// TIA Portal project "Project2" (V17)

(* hardware
DEVICE "S7-1500/ET200MP station_1"  S7-1500 station
   slot 0: "Rail_0"  Rack  6ES7 590-1***0-0AA0
   slot 1: "PLC_2"  CPU 1515-2 PN  6ES7 515-2AM00-0AB0  V1.8
      slot 3: "CPU display_1"  6ES7591-1BA00-0AA0
      slot 32768: "PROFINET interface_1"  X1
         slot 32769: "Port_1"  X1 P1
         slot 32770: "Port_2"  X1 P2
      slot 33024: "PROFINET interface_2"  X2
         slot 33025: "Port_1"  X2 P1
*)

// ===== PLC "PLC_2"  CPU 1515-2 PN =====

// folder: UDT/S2-Process Function Unit

TYPE "UDT_IS28xx_To_Plc"
   STRUCT
      iTriggerReady : Bool;   // This bit indicates when an In-Sight device can accept a new trigger via the Trigger bit. This field is true when the Trigger Enable bit is set, and the vision system is not currently acquiring an image.
      iTriggerAck : Bool;   // This bit indicates when an In-Sight device is successfully triggered via the Trigger bit. The Trigger Acknowledge bit stays set until the Trigger bit is cleared.
      iExposureComplete : Bool;   // This bit is set when the vision system image sensor is no longer exposed to light. It is used to indicate that the part being inspected can be moved from under the vision system's field of view.
      iAcquisitionError : Bool;   // This bit is set when an In-Sight device fails to acquire an image for one of the following reasons:
      iOfflineReason_1 : Bool;   // OfflineReason_1
      iOfflineReason_2 : Bool;   // OfflineReason_2
      iOfflineReason_3 : Bool;   // OfflineReason_3
      iSystemOnline : Bool;   // This bit indicates that the In-Sight device is online and the $System.OnlineEnabled tag is True.
      iReserve_1 : Byte;   // Reserve1
      iAcquisitonID : Int;   // This ID increments on the completion of every acquisition, regardless of the trigger source, and can be used to synchronize an acquisition with its Inspection Result. The Acquisition ID is changed on the start of an acquisition. If the PLC is the trigger source, the Acquisition ID is set prior to setting the Trigger Acknowledge bit.
      iReserve_2 : Bool;   // Reserve2
      iInspectionComplete : Bool;   // This bit is toggled upon the completion of an inspection.
      iResultBufferOverRun : Bool;   // This bit is set when the Enable Results Buffer bit is set, and there are more results than the result queue can hold.
      iResultValid : Bool;   // This bit is set when the Inspected Image ID, Inspection Result Code and Inspection Results fields are valid. The bit is cleared when the Inspection Results Acknowledge bit is set.
      iCommandExecuted : Bool;   // This bit is set while a command execution is in progress.
      iCommandComplete : Bool;   // This bit is set when the command execution is completed, and cleared when the Execute Command bit has been cleare
      iCommandFailed : Bool;   // This bit is set on the completion of a command, if the command has failed to execute successfully, or if an unknown Command ID was set.
      iSetUserDataAck : Bool;   // This bit is set to acknowledge completion of the Set User Data command.
      iJobPass : Bool;   // This bit indicates the pass and/or fail state of the inspection.
      iReserve_3 : Bool;   // Reserve3
      iReserve_4 : Bool;   // Reserve4
      iReserve_5 : Bool;   // Reserve5
      iReserve_6 : Bool;   // Reserve6
      iReserve_7 : Bool;   // Reserve7
      iReserve_8 : Bool;   // Reserve8
      iError : Bool;   // This bit is set when an error has occurred, which is defined in the Error ID field.
      iErrorID : Int;   // See Error ID codes.
      iCurrentRunningJobID : Int;   // These bits indicate the pre-added number of the current job filename. A job ID is a 16 bit number from 0 to 65535, but the PLC function can only load job IDs between 0‑999.
      iCommandResultCode : Int;   // This field is used to indicate the reason a command failed to execute successfully (the code is specific to the command executed):
      iExternalSoftEventAck : Byte;   // The External Event Acknowledge will be generated after the associated script finishes its execution
      iInspectionResultData : Struct
         iInspectionID : Int;   // The acquisition ID associated with this set of results.
         iInspectionResultCode : Int;   // These bytes are used to pass the user-defined result code. The inspection result code is defined by the Result Code parameter of the WriteResultsBuffer function
         iInspectionResult : Array[1..60] of Byte;   // These bytes of the inspection tool results can be written to the currently enabled factory communication protocol via the WriteResultsBuffer function.
      END_STRUCT;
   END_STRUCT;
END_TYPE

TYPE "UDT_Plc_To_IS28xx"
   STRUCT
      qTriggerEnable : Bool;   // This field is set to enable triggering via the Trigger bit. Clear this bit to disable the network triggering mechanism
      qTrigger : Bool;   // Setting the Trigger bit will trigger an acquisition on the vision system. The Trigger Enable bit must also be set
      qClearExposureComplete : Bool;   // When this signal is held high, the Exposure Complete status will remain reset. Once this signal is set to low, the Exposure Complete status will be set to high on the next exposure completion.
      qReserve_1 : Bool;   // Reserve_1
      qReserve_2 : Bool;   // Reserve_2
      qReserve_3 : Bool;   // Reserve_3
      qReserve_4 : Bool;   // Reserve_4
      qSetOffline : Bool;   // When this bit is set, the In-Sight vision system is paused and the state of the $System.OnlineEnabledComm is false
      qBufferResultEnable : Bool;   // When this bit is set, the Inspection ID, Inspection Result and Inspection Results fields are held constant until the Inspection Results Acknowledge field has acknowledged them and been set. Up to 16 sets of results are held in the buffer. Each result must be explicitly acknowledged using the Inspection Results Acknowledge signal.
      qInspectionResultAck : Bool;   // When the Buffer Results Enable bit is set, the Inspection Results Acknowledge bit acknowledges that the PLC has received the Inspected Image ID, Inspection Result Code and Inspection Results data.
      qSetUserData : Bool;   // This bit is used to signal that new User Data is available to be read in the vision system. After latching the entire User Data area into a holding buffer, the vision system will indicate to the PLC that it has read the data, and it can start loading new data into the buffer, if required, by issuing the Set User Data Acknowledge signal.
      qExecuteCommand : Bool;   // When the Execute Command bit is set to high, the Command ID signal is read by the vision system and the associated command is executed. The signal must be held high until the Command Completed bit is set. Once the Command Completed bit is set, clearing the Execute Command bit also clears the Command Completed bit.
      qReserve_5 : Bool;   // Reserve_5
      qReserve_6 : Bool;   // Reserve_6
      qReserve_7 : Bool;   // Reserve_7
      qClearError : Bool;   // When this bit is set, it clears the Error and Error ID signals; the Clear Error bit need to be held high until the Error bit is cleared. If an error is queued, clearing this bit causes the Error and Error ID signals to be set to the next queued error code.
      qCommandID : Int;   // This field indicates the command that will be executed on the rising edge of the Execute Command bit. This signal should not be changed until the Command Completed bit has been set.
      qSoftControlInput : Byte;   // Setting the External Event allows the PLC to trigger an associated event in the Spreadsheet.
      qUserData : Array[1..60] of Byte;   // Data buffer which can be read into the spreadsheet using the ReadUserDataBuffer function. The buffer is written exactly as it appears in the PLC
   END_STRUCT;
END_TYPE

// folder: (top level)

FUNCTION_BLOCK "PR_CentreStand_Fix_Seq_V12_1026b5"   // FB1, LAD
{ S7_Optimized_Access := 'TRUE' }
VERSION : 0.1
   VAR_INPUT
      iAutoRunning : Bool;
      iFixClamp : Bool;
      iFixEmpty : Bool;
      iFixTrayPresent : Bool;
      iFixUnclamp : Bool;
      iR1DropOver : Bool;
      iR1PickOver : Bool;
      iR2OperationOver : Bool;
      iR2ServiceActivated : Bool;
      iReset_fault : Bool;
      iRobotOutofZone : Bool;
      iSstMode : Bool;
      iSstPB : Bool;
   END_VAR
   VAR_OUTPUT
      qFixClamp : Bool;
      qFixUnclamp : Bool;
      qR1ReadytoDropTray : Bool;
      qR1ReadytoPickTray : Bool;
      qR2OperationStart : Bool;
   END_VAR
   VAR_IN_OUT
      iqR2ServiceActive : Bool;
      iqR2ServiceCompleted : Bool;
   END_VAR
   VAR
      StateNo : Int;
      s138_WaitBothRbtOutAl : Bool;
      s138_WaitBothRbtOutAl_T1 : Bool;
      s138_WaitBothRbtOutAl_T2 : Bool;
      s139_FixEmpty : Bool;
      s139_FixEmpty_T1 : Bool;
      s140_FixTrayPrsntRec : Bool;
      s140_FixTrayPrsntRec_T1 : Bool;
      s140_FixTrayPrsntRec_T2 : Bool;
      s141_FixUnclampCmd : Bool;
      s141_FixUnclampCmd_T1 : Bool;
      s142_TrayRdyDropFix : Bool;
      s142_TrayRdyDropFix_T1 : Bool;
      s143_RbtDropFixChkTr : Bool;
      s143_RbtDropFixChkTr_T1 : Bool;
      s144_RbtOutAreaDrop : Bool;
      s144_RbtOutAreaDrop_T1 : Bool;
      s145_FixClamp : Bool;
      s145_FixClamp_T1 : Bool;
      s146_Rbt2AlloyOpOver : Bool;
      s146_Rbt2AlloyOpOver_T1 : Bool;
      s147_FixUnclmpCmdAft : Bool;
      s147_FixUnclmpCmdAft_T1 : Bool;
      s148_RdyPickTrayAftr : Bool;
      s148_RdyPickTrayAftr_T1 : Bool;
      s149_RbtPickTrayChkE : Bool;
      s149_RbtPickTrayChkE_T1 : Bool;
      s191_WaitRbt2OutArea : Bool;
      s191_WaitRbt2OutArea_T1 : Bool;
      sSst : Bool;
      sSstPulse : Bool;
      sSstRise : Bool;
      sStWtResetRel : Bool;
      sStWtResetRel_T1 : Bool;
   END_VAR
   VAR_TEMP
      c138_WaitBothRbtOutAl_T1 : Bool;
      c138_WaitBothRbtOutAl_T2 : Bool;
      c140_FixTrayPrsntRec_T1 : Bool;
      c140_FixTrayPrsntRec_T2 : Bool;
      tOne : Bool;
   END_VAR
   VAR_TEMP   // added for the SCL form of the ladder/FBD networks
      _w1 : Bool;
   END_VAR
BEGIN

REGION Network 1
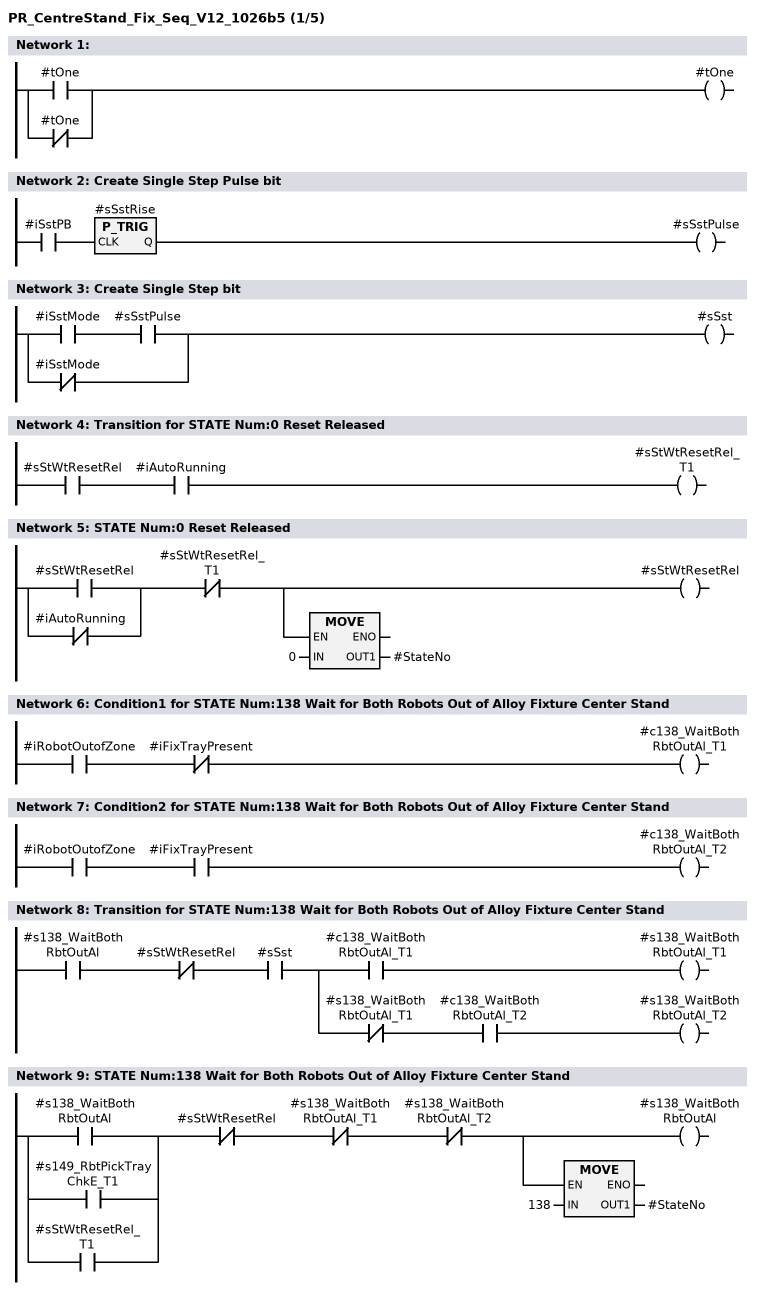
   RUNG wire#powerrail
      Contact( #tOne )
      wire#w1
      Coil( #tOne )
   END_RUNG
   RUNG wire#powerrail
      I_Contact( #tOne )
   END_RUNG wire#w1
   // the same network as SCL:
   #tOne := #tOne OR NOT #tOne;
END_REGION

REGION Network 2: Create Single Step Pulse bit
   RUNG wire#powerrail
      Contact( #iSstPB )
      P_Trig( #sSstRise )
      Coil( #sSstPulse )
   END_RUNG
   // the same network as SCL:
   #_w1 := #iSstPB AND NOT #sSstRise;   // rising edge
   #sSstRise := #iSstPB;
   #sSstPulse := #_w1;
END_REGION

REGION Network 3: Create Single Step bit
   RUNG wire#powerrail
      Contact( #iSstMode )
      Contact( #sSstPulse )
      wire#w1
      Coil( #sSst )
   END_RUNG
   RUNG wire#powerrail
      I_Contact( #iSstMode )
   END_RUNG wire#w1
   // the same network as SCL:
   #sSst := (#iSstMode AND #sSstPulse) OR NOT #iSstMode;
END_REGION

REGION Network 4: Transition for STATE Num:0 Reset Released
   RUNG wire#powerrail
      Contact( #sStWtResetRel )
      Contact( #iAutoRunning )
      Coil( #sStWtResetRel_T1 )
   END_RUNG
   // the same network as SCL:
   #sStWtResetRel_T1 := #sStWtResetRel AND #iAutoRunning;
END_REGION

REGION Network 5: STATE Num:0 Reset Released
   RUNG wire#powerrail
      Contact( #sStWtResetRel )
      wire#w1
      I_Contact( #sStWtResetRel_T1 )
      wire#w2
      Coil( #sStWtResetRel )
   END_RUNG
   RUNG wire#powerrail
      I_Contact( #iAutoRunning )
   END_RUNG wire#w1
   RUNG wire#w2
      { S7_GenerateENO := "TRUE" } Move(in := 0, out1 => #StateNo)
   END_RUNG
   // the same network as SCL:
   #sStWtResetRel := (#sStWtResetRel OR NOT #iAutoRunning) AND NOT #sStWtResetRel_T1;
   IF #sStWtResetRel THEN #StateNo := 0; END_IF;
END_REGION

REGION Network 6: Condition1 for STATE Num:138 Wait for Both Robots Out of Alloy Fixture Center Stand
   RUNG wire#powerrail
      Contact( #iRobotOutofZone )
      I_Contact( #iFixTrayPresent )
      Coil( #c138_WaitBothRbtOutAl_T1 )
   END_RUNG
   // the same network as SCL:
   #c138_WaitBothRbtOutAl_T1 := #iRobotOutofZone AND NOT #iFixTrayPresent;
END_REGION

REGION Network 7: Condition2 for STATE Num:138 Wait for Both Robots Out of Alloy Fixture Center Stand
   RUNG wire#powerrail
      Contact( #iRobotOutofZone )
      Contact( #iFixTrayPresent )
      Coil( #c138_WaitBothRbtOutAl_T2 )
   END_RUNG
   // the same network as SCL:
   #c138_WaitBothRbtOutAl_T2 := #iRobotOutofZone AND #iFixTrayPresent;
END_REGION

REGION Network 8: Transition for STATE Num:138 Wait for Both Robots Out of Alloy Fixture Center Stand
   RUNG wire#powerrail
      Contact( #s138_WaitBothRbtOutAl )
      I_Contact( #sStWtResetRel )
      Contact( #sSst )
      wire#w1
      Contact( #c138_WaitBothRbtOutAl_T1 )
      Coil( #s138_WaitBothRbtOutAl_T1 )
   END_RUNG
   RUNG wire#w1
      I_Contact( #s138_WaitBothRbtOutAl_T1 )
      Contact( #c138_WaitBothRbtOutAl_T2 )
      Coil( #s138_WaitBothRbtOutAl_T2 )
   END_RUNG
   // the same network as SCL:
   #_w1 := #s138_WaitBothRbtOutAl AND NOT #sStWtResetRel AND #sSst;
   #s138_WaitBothRbtOutAl_T1 := #_w1 AND #c138_WaitBothRbtOutAl_T1;
   #s138_WaitBothRbtOutAl_T2 := #_w1 AND NOT #s138_WaitBothRbtOutAl_T1 AND #c138_WaitBothRbtOutAl_T2;
END_REGION

REGION Network 9: STATE Num:138 Wait for Both Robots Out of Alloy Fixture Center Stand
   RUNG wire#powerrail
      Contact( #s138_WaitBothRbtOutAl )
      wire#w1
      I_Contact( #sStWtResetRel )
      I_Contact( #s138_WaitBothRbtOutAl_T1 )
      I_Contact( #s138_WaitBothRbtOutAl_T2 )
      wire#w2
      Coil( #s138_WaitBothRbtOutAl )
   END_RUNG
   RUNG wire#powerrail
      Contact( #s149_RbtPickTrayChkE_T1 )
   END_RUNG wire#w1
   RUNG wire#powerrail
      Contact( #sStWtResetRel_T1 )
   END_RUNG wire#w1
   RUNG wire#w2
      { S7_GenerateENO := "TRUE" } Move(in := 138, out1 => #StateNo)
   END_RUNG
   // the same network as SCL:
   #s138_WaitBothRbtOutAl := (#s138_WaitBothRbtOutAl OR #s149_RbtPickTrayChkE_T1 OR #sStWtResetRel_T1) AND NOT #sStWtResetRel AND NOT #s138_WaitBothRbtOutAl_T1 AND NOT #s138_WaitBothRbtOutAl_T2;
   IF #s138_WaitBothRbtOutAl THEN #StateNo := 138; END_IF;
END_REGION

REGION Network 10: Transition for STATE Num:139 Fix Empty
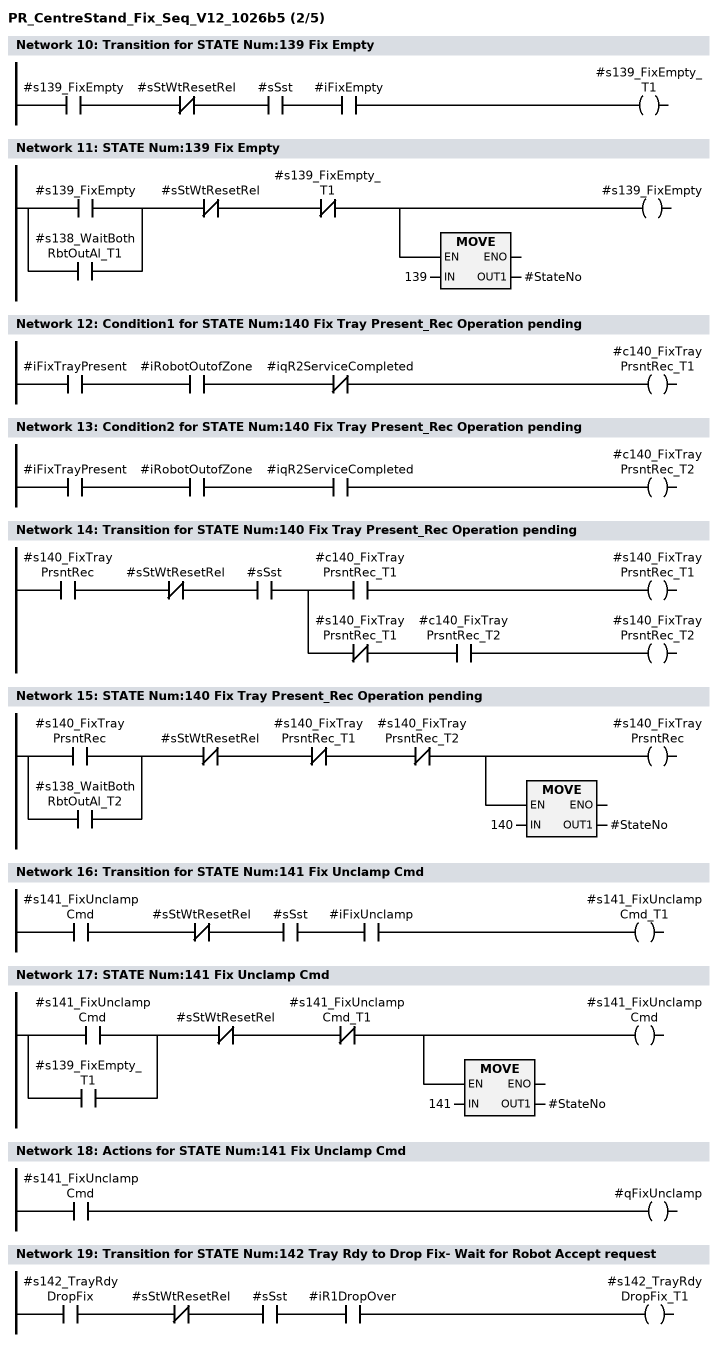
   RUNG wire#powerrail
      Contact( #s139_FixEmpty )
      I_Contact( #sStWtResetRel )
      Contact( #sSst )
      Contact( #iFixEmpty )
      Coil( #s139_FixEmpty_T1 )
   END_RUNG
   // the same network as SCL:
   #s139_FixEmpty_T1 := #s139_FixEmpty AND NOT #sStWtResetRel AND #sSst AND #iFixEmpty;
END_REGION

REGION Network 11: STATE Num:139 Fix Empty
   RUNG wire#powerrail
      Contact( #s139_FixEmpty )
      wire#w1
      I_Contact( #sStWtResetRel )
      I_Contact( #s139_FixEmpty_T1 )
      wire#w2
      Coil( #s139_FixEmpty )
   END_RUNG
   RUNG wire#powerrail
      Contact( #s138_WaitBothRbtOutAl_T1 )
   END_RUNG wire#w1
   RUNG wire#w2
      { S7_GenerateENO := "TRUE" } Move(in := 139, out1 => #StateNo)
   END_RUNG
   // the same network as SCL:
   #s139_FixEmpty := (#s139_FixEmpty OR #s138_WaitBothRbtOutAl_T1) AND NOT #sStWtResetRel AND NOT #s139_FixEmpty_T1;
   IF #s139_FixEmpty THEN #StateNo := 139; END_IF;
END_REGION

REGION Network 12: Condition1 for STATE Num:140 Fix Tray Present_Rec Operation pending
   RUNG wire#powerrail
      Contact( #iFixTrayPresent )
      Contact( #iRobotOutofZone )
      I_Contact( #iqR2ServiceCompleted )
      Coil( #c140_FixTrayPrsntRec_T1 )
   END_RUNG
   // the same network as SCL:
   #c140_FixTrayPrsntRec_T1 := #iFixTrayPresent AND #iRobotOutofZone AND NOT #iqR2ServiceCompleted;
END_REGION

REGION Network 13: Condition2 for STATE Num:140 Fix Tray Present_Rec Operation pending
   RUNG wire#powerrail
      Contact( #iFixTrayPresent )
      Contact( #iRobotOutofZone )
      Contact( #iqR2ServiceCompleted )
      Coil( #c140_FixTrayPrsntRec_T2 )
   END_RUNG
   // the same network as SCL:
   #c140_FixTrayPrsntRec_T2 := #iFixTrayPresent AND #iRobotOutofZone AND #iqR2ServiceCompleted;
END_REGION

REGION Network 14: Transition for STATE Num:140 Fix Tray Present_Rec Operation pending
   RUNG wire#powerrail
      Contact( #s140_FixTrayPrsntRec )
      I_Contact( #sStWtResetRel )
      Contact( #sSst )
      wire#w1
      Contact( #c140_FixTrayPrsntRec_T1 )
      Coil( #s140_FixTrayPrsntRec_T1 )
   END_RUNG
   RUNG wire#w1
      I_Contact( #s140_FixTrayPrsntRec_T1 )
      Contact( #c140_FixTrayPrsntRec_T2 )
      Coil( #s140_FixTrayPrsntRec_T2 )
   END_RUNG
   // the same network as SCL:
   #_w1 := #s140_FixTrayPrsntRec AND NOT #sStWtResetRel AND #sSst;
   #s140_FixTrayPrsntRec_T1 := #_w1 AND #c140_FixTrayPrsntRec_T1;
   #s140_FixTrayPrsntRec_T2 := #_w1 AND NOT #s140_FixTrayPrsntRec_T1 AND #c140_FixTrayPrsntRec_T2;
END_REGION

REGION Network 15: STATE Num:140 Fix Tray Present_Rec Operation pending
   RUNG wire#powerrail
      Contact( #s140_FixTrayPrsntRec )
      wire#w1
      I_Contact( #sStWtResetRel )
      I_Contact( #s140_FixTrayPrsntRec_T1 )
      I_Contact( #s140_FixTrayPrsntRec_T2 )
      wire#w2
      Coil( #s140_FixTrayPrsntRec )
   END_RUNG
   RUNG wire#powerrail
      Contact( #s138_WaitBothRbtOutAl_T2 )
   END_RUNG wire#w1
   RUNG wire#w2
      { S7_GenerateENO := "TRUE" } Move(in := 140, out1 => #StateNo)
   END_RUNG
   // the same network as SCL:
   #s140_FixTrayPrsntRec := (#s140_FixTrayPrsntRec OR #s138_WaitBothRbtOutAl_T2) AND NOT #sStWtResetRel AND NOT #s140_FixTrayPrsntRec_T1 AND NOT #s140_FixTrayPrsntRec_T2;
   IF #s140_FixTrayPrsntRec THEN #StateNo := 140; END_IF;
END_REGION

REGION Network 16: Transition for STATE Num:141 Fix Unclamp Cmd
   RUNG wire#powerrail
      Contact( #s141_FixUnclampCmd )
      I_Contact( #sStWtResetRel )
      Contact( #sSst )
      Contact( #iFixUnclamp )
      Coil( #s141_FixUnclampCmd_T1 )
   END_RUNG
   // the same network as SCL:
   #s141_FixUnclampCmd_T1 := #s141_FixUnclampCmd AND NOT #sStWtResetRel AND #sSst AND #iFixUnclamp;
END_REGION

REGION Network 17: STATE Num:141 Fix Unclamp Cmd
   RUNG wire#powerrail
      Contact( #s141_FixUnclampCmd )
      wire#w1
      I_Contact( #sStWtResetRel )
      I_Contact( #s141_FixUnclampCmd_T1 )
      wire#w2
      Coil( #s141_FixUnclampCmd )
   END_RUNG
   RUNG wire#powerrail
      Contact( #s139_FixEmpty_T1 )
   END_RUNG wire#w1
   RUNG wire#w2
      { S7_GenerateENO := "TRUE" } Move(in := 141, out1 => #StateNo)
   END_RUNG
   // the same network as SCL:
   #s141_FixUnclampCmd := (#s141_FixUnclampCmd OR #s139_FixEmpty_T1) AND NOT #sStWtResetRel AND NOT #s141_FixUnclampCmd_T1;
   IF #s141_FixUnclampCmd THEN #StateNo := 141; END_IF;
END_REGION

REGION Network 18: Actions for STATE Num:141 Fix Unclamp Cmd
   RUNG wire#powerrail
      Contact( #s141_FixUnclampCmd )
      Coil( #qFixUnclamp )
   END_RUNG
   // the same network as SCL:
   #qFixUnclamp := #s141_FixUnclampCmd;
END_REGION

REGION Network 19: Transition for STATE Num:142 Tray Rdy to Drop Fix- Wait for Robot Accept request
   RUNG wire#powerrail
      Contact( #s142_TrayRdyDropFix )
      I_Contact( #sStWtResetRel )
      Contact( #sSst )
      Contact( #iR1DropOver )
      Coil( #s142_TrayRdyDropFix_T1 )
   END_RUNG
   // the same network as SCL:
   #s142_TrayRdyDropFix_T1 := #s142_TrayRdyDropFix AND NOT #sStWtResetRel AND #sSst AND #iR1DropOver;
END_REGION

REGION Network 20: STATE Num:142 Tray Rdy to Drop Fix- Wait for Robot Accept request
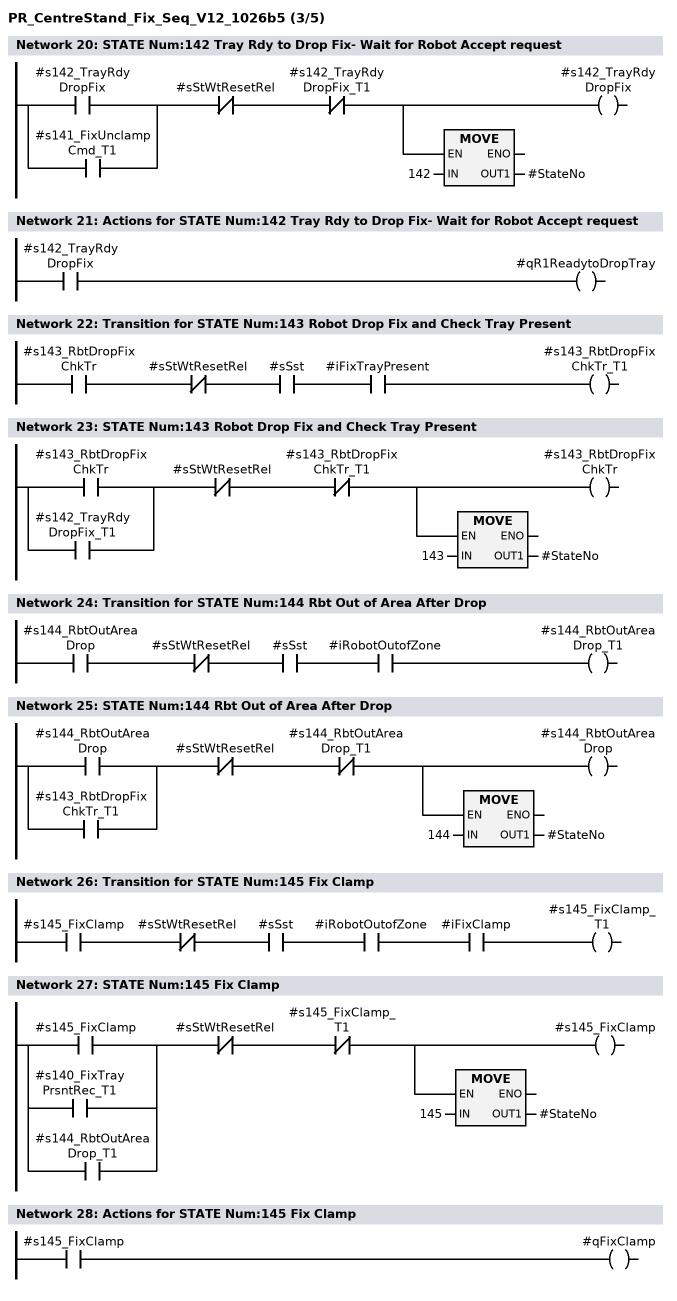
   RUNG wire#powerrail
      Contact( #s142_TrayRdyDropFix )
      wire#w1
      I_Contact( #sStWtResetRel )
      I_Contact( #s142_TrayRdyDropFix_T1 )
      wire#w2
      Coil( #s142_TrayRdyDropFix )
   END_RUNG
   RUNG wire#powerrail
      Contact( #s141_FixUnclampCmd_T1 )
   END_RUNG wire#w1
   RUNG wire#w2
      { S7_GenerateENO := "TRUE" } Move(in := 142, out1 => #StateNo)
   END_RUNG
   // the same network as SCL:
   #s142_TrayRdyDropFix := (#s142_TrayRdyDropFix OR #s141_FixUnclampCmd_T1) AND NOT #sStWtResetRel AND NOT #s142_TrayRdyDropFix_T1;
   IF #s142_TrayRdyDropFix THEN #StateNo := 142; END_IF;
END_REGION

REGION Network 21: Actions for STATE Num:142 Tray Rdy to Drop Fix- Wait for Robot Accept request
   RUNG wire#powerrail
      Contact( #s142_TrayRdyDropFix )
      Coil( #qR1ReadytoDropTray )
   END_RUNG
   // the same network as SCL:
   #qR1ReadytoDropTray := #s142_TrayRdyDropFix;
END_REGION

REGION Network 22: Transition for STATE Num:143 Robot Drop Fix and Check Tray Present
   RUNG wire#powerrail
      Contact( #s143_RbtDropFixChkTr )
      I_Contact( #sStWtResetRel )
      Contact( #sSst )
      Contact( #iFixTrayPresent )
      Coil( #s143_RbtDropFixChkTr_T1 )
   END_RUNG
   // the same network as SCL:
   #s143_RbtDropFixChkTr_T1 := #s143_RbtDropFixChkTr AND NOT #sStWtResetRel AND #sSst AND #iFixTrayPresent;
END_REGION

REGION Network 23: STATE Num:143 Robot Drop Fix and Check Tray Present
   RUNG wire#powerrail
      Contact( #s143_RbtDropFixChkTr )
      wire#w1
      I_Contact( #sStWtResetRel )
      I_Contact( #s143_RbtDropFixChkTr_T1 )
      wire#w2
      Coil( #s143_RbtDropFixChkTr )
   END_RUNG
   RUNG wire#powerrail
      Contact( #s142_TrayRdyDropFix_T1 )
   END_RUNG wire#w1
   RUNG wire#w2
      { S7_GenerateENO := "TRUE" } Move(in := 143, out1 => #StateNo)
   END_RUNG
   // the same network as SCL:
   #s143_RbtDropFixChkTr := (#s143_RbtDropFixChkTr OR #s142_TrayRdyDropFix_T1) AND NOT #sStWtResetRel AND NOT #s143_RbtDropFixChkTr_T1;
   IF #s143_RbtDropFixChkTr THEN #StateNo := 143; END_IF;
END_REGION

REGION Network 24: Transition for STATE Num:144 Rbt Out of Area After Drop
   RUNG wire#powerrail
      Contact( #s144_RbtOutAreaDrop )
      I_Contact( #sStWtResetRel )
      Contact( #sSst )
      Contact( #iRobotOutofZone )
      Coil( #s144_RbtOutAreaDrop_T1 )
   END_RUNG
   // the same network as SCL:
   #s144_RbtOutAreaDrop_T1 := #s144_RbtOutAreaDrop AND NOT #sStWtResetRel AND #sSst AND #iRobotOutofZone;
END_REGION

REGION Network 25: STATE Num:144 Rbt Out of Area After Drop
   RUNG wire#powerrail
      Contact( #s144_RbtOutAreaDrop )
      wire#w1
      I_Contact( #sStWtResetRel )
      I_Contact( #s144_RbtOutAreaDrop_T1 )
      wire#w2
      Coil( #s144_RbtOutAreaDrop )
   END_RUNG
   RUNG wire#powerrail
      Contact( #s143_RbtDropFixChkTr_T1 )
   END_RUNG wire#w1
   RUNG wire#w2
      { S7_GenerateENO := "TRUE" } Move(in := 144, out1 => #StateNo)
   END_RUNG
   // the same network as SCL:
   #s144_RbtOutAreaDrop := (#s144_RbtOutAreaDrop OR #s143_RbtDropFixChkTr_T1) AND NOT #sStWtResetRel AND NOT #s144_RbtOutAreaDrop_T1;
   IF #s144_RbtOutAreaDrop THEN #StateNo := 144; END_IF;
END_REGION

REGION Network 26: Transition for STATE Num:145 Fix Clamp
   RUNG wire#powerrail
      Contact( #s145_FixClamp )
      I_Contact( #sStWtResetRel )
      Contact( #sSst )
      Contact( #iRobotOutofZone )
      Contact( #iFixClamp )
      Coil( #s145_FixClamp_T1 )
   END_RUNG
   // the same network as SCL:
   #s145_FixClamp_T1 := #s145_FixClamp AND NOT #sStWtResetRel AND #sSst AND #iRobotOutofZone AND #iFixClamp;
END_REGION

REGION Network 27: STATE Num:145 Fix Clamp
   RUNG wire#powerrail
      Contact( #s145_FixClamp )
      wire#w1
      I_Contact( #sStWtResetRel )
      I_Contact( #s145_FixClamp_T1 )
      wire#w2
      Coil( #s145_FixClamp )
   END_RUNG
   RUNG wire#powerrail
      Contact( #s140_FixTrayPrsntRec_T1 )
   END_RUNG wire#w1
   RUNG wire#powerrail
      Contact( #s144_RbtOutAreaDrop_T1 )
   END_RUNG wire#w1
   RUNG wire#w2
      { S7_GenerateENO := "TRUE" } Move(in := 145, out1 => #StateNo)
   END_RUNG
   // the same network as SCL:
   #s145_FixClamp := (#s145_FixClamp OR #s140_FixTrayPrsntRec_T1 OR #s144_RbtOutAreaDrop_T1) AND NOT #sStWtResetRel AND NOT #s145_FixClamp_T1;
   IF #s145_FixClamp THEN #StateNo := 145; END_IF;
END_REGION

REGION Network 28: Actions for STATE Num:145 Fix Clamp
   RUNG wire#powerrail
      Contact( #s145_FixClamp )
      Coil( #qFixClamp )
   END_RUNG
   // the same network as SCL:
   #qFixClamp := #s145_FixClamp;
END_REGION

REGION Network 29: Transition for STATE Num:146 Robot-2 All Alloys Pick Or Drop Operation over
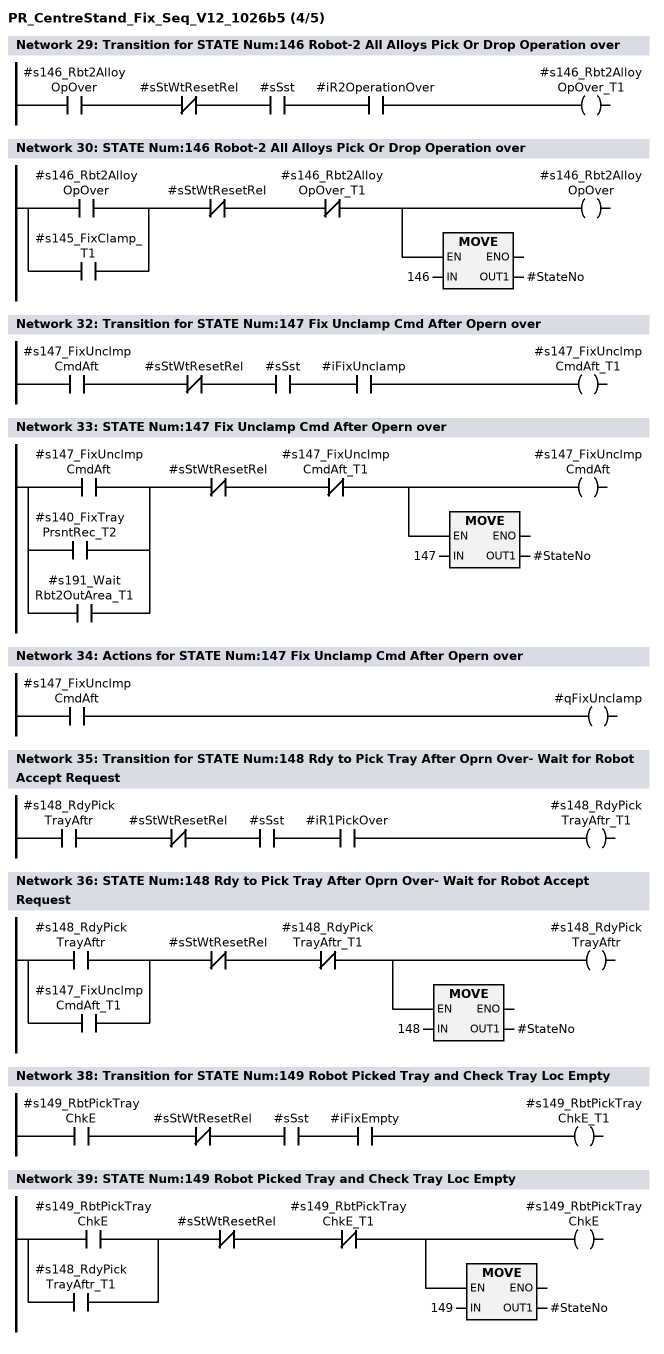
   RUNG wire#powerrail
      Contact( #s146_Rbt2AlloyOpOver )
      I_Contact( #sStWtResetRel )
      Contact( #sSst )
      Contact( #iR2OperationOver )
      Coil( #s146_Rbt2AlloyOpOver_T1 )
   END_RUNG
   // the same network as SCL:
   #s146_Rbt2AlloyOpOver_T1 := #s146_Rbt2AlloyOpOver AND NOT #sStWtResetRel AND #sSst AND #iR2OperationOver;
END_REGION

REGION Network 30: STATE Num:146 Robot-2 All Alloys Pick Or Drop Operation over
   RUNG wire#powerrail
      Contact( #s146_Rbt2AlloyOpOver )
      wire#w1
      I_Contact( #sStWtResetRel )
      I_Contact( #s146_Rbt2AlloyOpOver_T1 )
      wire#w2
      Coil( #s146_Rbt2AlloyOpOver )
   END_RUNG
   RUNG wire#powerrail
      Contact( #s145_FixClamp_T1 )
   END_RUNG wire#w1
   RUNG wire#w2
      { S7_GenerateENO := "TRUE" } Move(in := 146, out1 => #StateNo)
   END_RUNG
   // the same network as SCL:
   #s146_Rbt2AlloyOpOver := (#s146_Rbt2AlloyOpOver OR #s145_FixClamp_T1) AND NOT #sStWtResetRel AND NOT #s146_Rbt2AlloyOpOver_T1;
   IF #s146_Rbt2AlloyOpOver THEN #StateNo := 146; END_IF;
END_REGION

REGION Network 31 (STL): Actions for STATE Num:146 Robot-2 All Alloys Pick Or Drop Operation over
         A     #s146_Rbt2AlloyOpOver;
         =     #qR2OperationStart;
         A     #s146_Rbt2AlloyOpOver;
         A     #iR2ServiceActivated;
         S     #iqR2ServiceActive;
         A     #s146_Rbt2AlloyOpOver;
         A     #iR2OperationOver;
         A     #iqR2ServiceActive;
         R     #iqR2ServiceActive;
END_REGION

REGION Network 32: Transition for STATE Num:147 Fix Unclamp Cmd After Opern over
   RUNG wire#powerrail
      Contact( #s147_FixUnclmpCmdAft )
      I_Contact( #sStWtResetRel )
      Contact( #sSst )
      Contact( #iFixUnclamp )
      Coil( #s147_FixUnclmpCmdAft_T1 )
   END_RUNG
   // the same network as SCL:
   #s147_FixUnclmpCmdAft_T1 := #s147_FixUnclmpCmdAft AND NOT #sStWtResetRel AND #sSst AND #iFixUnclamp;
END_REGION

REGION Network 33: STATE Num:147 Fix Unclamp Cmd After Opern over
   RUNG wire#powerrail
      Contact( #s147_FixUnclmpCmdAft )
      wire#w1
      I_Contact( #sStWtResetRel )
      I_Contact( #s147_FixUnclmpCmdAft_T1 )
      wire#w2
      Coil( #s147_FixUnclmpCmdAft )
   END_RUNG
   RUNG wire#powerrail
      Contact( #s140_FixTrayPrsntRec_T2 )
   END_RUNG wire#w1
   RUNG wire#powerrail
      Contact( #s191_WaitRbt2OutArea_T1 )
   END_RUNG wire#w1
   RUNG wire#w2
      { S7_GenerateENO := "TRUE" } Move(in := 147, out1 => #StateNo)
   END_RUNG
   // the same network as SCL:
   #s147_FixUnclmpCmdAft := (#s147_FixUnclmpCmdAft OR #s140_FixTrayPrsntRec_T2 OR #s191_WaitRbt2OutArea_T1) AND NOT #sStWtResetRel AND NOT #s147_FixUnclmpCmdAft_T1;
   IF #s147_FixUnclmpCmdAft THEN #StateNo := 147; END_IF;
END_REGION

REGION Network 34: Actions for STATE Num:147 Fix Unclamp Cmd After Opern over
   RUNG wire#powerrail
      Contact( #s147_FixUnclmpCmdAft )
      Coil( #qFixUnclamp )
   END_RUNG
   // the same network as SCL:
   #qFixUnclamp := #s147_FixUnclmpCmdAft;
END_REGION

REGION Network 35: Transition for STATE Num:148 Rdy to Pick Tray After Oprn Over- Wait for Robot Accept Request
   RUNG wire#powerrail
      Contact( #s148_RdyPickTrayAftr )
      I_Contact( #sStWtResetRel )
      Contact( #sSst )
      Contact( #iR1PickOver )
      Coil( #s148_RdyPickTrayAftr_T1 )
   END_RUNG
   // the same network as SCL:
   #s148_RdyPickTrayAftr_T1 := #s148_RdyPickTrayAftr AND NOT #sStWtResetRel AND #sSst AND #iR1PickOver;
END_REGION

REGION Network 36: STATE Num:148 Rdy to Pick Tray After Oprn Over- Wait for Robot Accept Request
   RUNG wire#powerrail
      Contact( #s148_RdyPickTrayAftr )
      wire#w1
      I_Contact( #sStWtResetRel )
      I_Contact( #s148_RdyPickTrayAftr_T1 )
      wire#w2
      Coil( #s148_RdyPickTrayAftr )
   END_RUNG
   RUNG wire#powerrail
      Contact( #s147_FixUnclmpCmdAft_T1 )
   END_RUNG wire#w1
   RUNG wire#w2
      { S7_GenerateENO := "TRUE" } Move(in := 148, out1 => #StateNo)
   END_RUNG
   // the same network as SCL:
   #s148_RdyPickTrayAftr := (#s148_RdyPickTrayAftr OR #s147_FixUnclmpCmdAft_T1) AND NOT #sStWtResetRel AND NOT #s148_RdyPickTrayAftr_T1;
   IF #s148_RdyPickTrayAftr THEN #StateNo := 148; END_IF;
END_REGION

REGION Network 37 (STL): Actions for STATE Num:148 Rdy to Pick Tray After Oprn Over- Wait for Robot Accept Request
         A     #s148_RdyPickTrayAftr;
         =     #qR1ReadytoPickTray;
         A     #s148_RdyPickTrayAftr;
         A     #iR1PickOver;
         R     #iqR2ServiceCompleted;
END_REGION

REGION Network 38: Transition for STATE Num:149 Robot Picked Tray and Check Tray Loc Empty
   RUNG wire#powerrail
      Contact( #s149_RbtPickTrayChkE )
      I_Contact( #sStWtResetRel )
      Contact( #sSst )
      Contact( #iFixEmpty )
      Coil( #s149_RbtPickTrayChkE_T1 )
   END_RUNG
   // the same network as SCL:
   #s149_RbtPickTrayChkE_T1 := #s149_RbtPickTrayChkE AND NOT #sStWtResetRel AND #sSst AND #iFixEmpty;
END_REGION

REGION Network 39: STATE Num:149 Robot Picked Tray and Check Tray Loc Empty
   RUNG wire#powerrail
      Contact( #s149_RbtPickTrayChkE )
      wire#w1
      I_Contact( #sStWtResetRel )
      I_Contact( #s149_RbtPickTrayChkE_T1 )
      wire#w2
      Coil( #s149_RbtPickTrayChkE )
   END_RUNG
   RUNG wire#powerrail
      Contact( #s148_RdyPickTrayAftr_T1 )
   END_RUNG wire#w1
   RUNG wire#w2
      { S7_GenerateENO := "TRUE" } Move(in := 149, out1 => #StateNo)
   END_RUNG
   // the same network as SCL:
   #s149_RbtPickTrayChkE := (#s149_RbtPickTrayChkE OR #s148_RdyPickTrayAftr_T1) AND NOT #sStWtResetRel AND NOT #s149_RbtPickTrayChkE_T1;
   IF #s149_RbtPickTrayChkE THEN #StateNo := 149; END_IF;
END_REGION

REGION Network 40: Actions for STATE Num:149 Robot Picked Tray and Check Tray Loc Empty
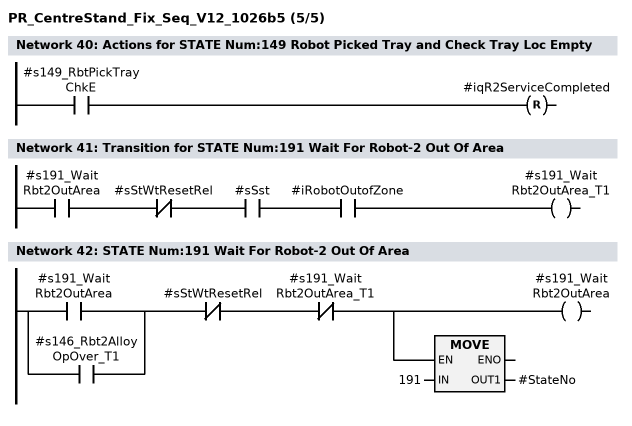
   RUNG wire#powerrail
      Contact( #s149_RbtPickTrayChkE )
      R_Coil( #iqR2ServiceCompleted )
   END_RUNG
   // the same network as SCL:
   IF #s149_RbtPickTrayChkE THEN #iqR2ServiceCompleted := FALSE; END_IF;
END_REGION

REGION Network 41: Transition for STATE Num:191 Wait For Robot-2 Out Of Area
   RUNG wire#powerrail
      Contact( #s191_WaitRbt2OutArea )
      I_Contact( #sStWtResetRel )
      Contact( #sSst )
      Contact( #iRobotOutofZone )
      Coil( #s191_WaitRbt2OutArea_T1 )
   END_RUNG
   // the same network as SCL:
   #s191_WaitRbt2OutArea_T1 := #s191_WaitRbt2OutArea AND NOT #sStWtResetRel AND #sSst AND #iRobotOutofZone;
END_REGION

REGION Network 42: STATE Num:191 Wait For Robot-2 Out Of Area
   RUNG wire#powerrail
      Contact( #s191_WaitRbt2OutArea )
      wire#w1
      I_Contact( #sStWtResetRel )
      I_Contact( #s191_WaitRbt2OutArea_T1 )
      wire#w2
      Coil( #s191_WaitRbt2OutArea )
   END_RUNG
   RUNG wire#powerrail
      Contact( #s146_Rbt2AlloyOpOver_T1 )
   END_RUNG wire#w1
   RUNG wire#w2
      { S7_GenerateENO := "TRUE" } Move(in := 191, out1 => #StateNo)
   END_RUNG
   // the same network as SCL:
   #s191_WaitRbt2OutArea := (#s191_WaitRbt2OutArea OR #s146_Rbt2AlloyOpOver_T1) AND NOT #sStWtResetRel AND NOT #s191_WaitRbt2OutArea_T1;
   IF #s191_WaitRbt2OutArea THEN #StateNo := 191; END_IF;
END_REGION
END_FUNCTION_BLOCK

FUNCTION_BLOCK "FB_CentreStand_Fix_Seq_2"   // FB1, LAD
{ S7_Optimized_Access := 'TRUE' }
VERSION : 0.1
   VAR_INPUT
      iAutoRunning : Bool;
      iFixClamp : Bool;
      iFixEmpty : Bool;
      iFixTrayPresent : Bool;
      iFixUnclamp : Bool;
      iR1DropOver : Bool;
      iR1PickOver : Bool;
      iR2OperationOver : Bool;
      iR2ServiceActivated : Bool;
      iR2ServiceCompleted : Bool;
      iReset_fault : Bool;
      iRobotOutofZone : Bool;
      iSstMode : Bool;
      iSstPB : Bool;
   END_VAR
   VAR_OUTPUT
      qFixClamp : Bool;
      qFixUnclamp : Bool;
      qR1ReadytoDropTray : Bool;
      qR1ReadytoPickTray : Bool;
      qR2OperationStart : Bool;
   END_VAR
   VAR_IN_OUT
      iqR2ServiceActive : Bool;
      iqR2ServiceCompleted : Bool;
   END_VAR
   VAR
      StateNo : Int;
      s138_WaitBothRbtOutAl : Bool;
      s138_WaitBothRbtOutAl_T1 : Bool;
      s138_WaitBothRbtOutAl_T2 : Bool;
      s139_FixEmpty : Bool;
      s139_FixEmpty_T1 : Bool;
      s140_FixTrayPrsntRec : Bool;
      s140_FixTrayPrsntRec_T1 : Bool;
      s140_FixTrayPrsntRec_T2 : Bool;
      s141_FixUnclampCmd : Bool;
      s141_FixUnclampCmd_T1 : Bool;
      s142_TrayRdyDropFix : Bool;
      s142_TrayRdyDropFix_T1 : Bool;
      s143_RbtDropFixChkTr : Bool;
      s143_RbtDropFixChkTr_T1 : Bool;
      s144_RbtOutAreaDrop : Bool;
      s144_RbtOutAreaDrop_T1 : Bool;
      s145_FixClamp : Bool;
      s145_FixClamp_T1 : Bool;
      s146_Rbt2AlloyOpOver : Bool;
      s146_Rbt2AlloyOpOver_T1 : Bool;
      s147_FixUnclmpCmdOvr : Bool;
      s147_FixUnclmpCmdOvr_T1 : Bool;
      s148_RdyPickTrayWait : Bool;
      s148_RdyPickTrayWait_T1 : Bool;
      s149_RbtPickTrayChkEm : Bool;
      s149_RbtPickTrayChkEm_T1 : Bool;
      s191_WaitRbt2OutArea : Bool;
      s191_WaitRbt2OutArea_T1 : Bool;
      sSst : Bool;
      sSstPulse : Bool;
      sSstRise : Bool;
      sStWtResetRel : Bool;
      sStWtResetRel_T1 : Bool;
   END_VAR
   VAR_TEMP
      tOne : Bool;
   END_VAR
   VAR_TEMP   // added for the SCL form of the ladder/FBD networks
      _w1 : Bool;
   END_VAR
BEGIN

REGION Network 1
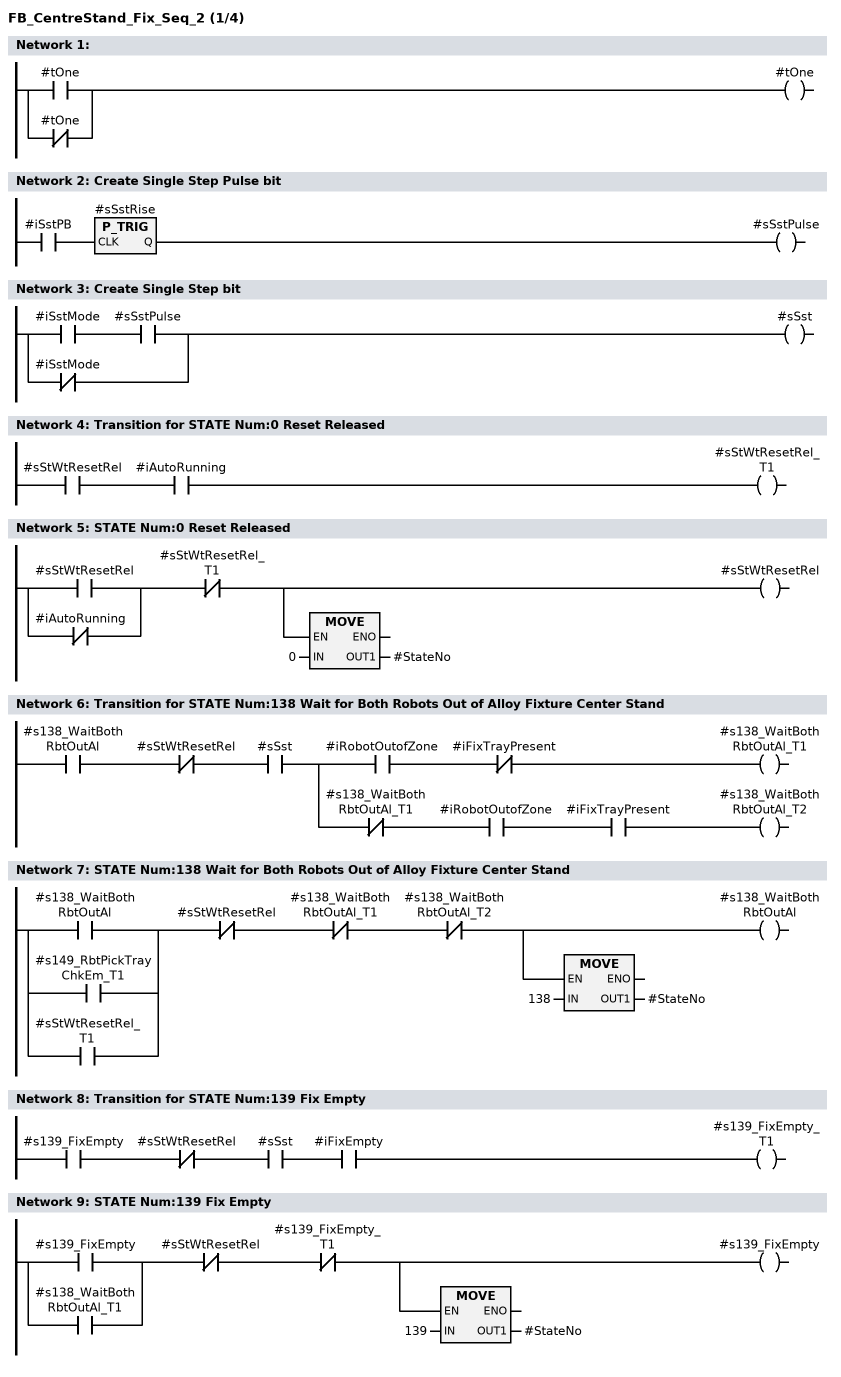
   RUNG wire#powerrail
      Contact( #tOne )
      wire#w1
      Coil( #tOne )
   END_RUNG
   RUNG wire#powerrail
      I_Contact( #tOne )
   END_RUNG wire#w1
   // the same network as SCL:
   #tOne := #tOne OR NOT #tOne;
END_REGION

REGION Network 2: Create Single Step Pulse bit
   RUNG wire#powerrail
      Contact( #iSstPB )
      P_Trig( #sSstRise )
      Coil( #sSstPulse )
   END_RUNG
   // the same network as SCL:
   #_w1 := #iSstPB AND NOT #sSstRise;   // rising edge
   #sSstRise := #iSstPB;
   #sSstPulse := #_w1;
END_REGION

REGION Network 3: Create Single Step bit
   RUNG wire#powerrail
      Contact( #iSstMode )
      Contact( #sSstPulse )
      wire#w1
      Coil( #sSst )
   END_RUNG
   RUNG wire#powerrail
      I_Contact( #iSstMode )
   END_RUNG wire#w1
   // the same network as SCL:
   #sSst := (#iSstMode AND #sSstPulse) OR NOT #iSstMode;
END_REGION

REGION Network 4: Transition for STATE Num:0 Reset Released
   RUNG wire#powerrail
      Contact( #sStWtResetRel )
      Contact( #iAutoRunning )
      Coil( #sStWtResetRel_T1 )
   END_RUNG
   // the same network as SCL:
   #sStWtResetRel_T1 := #sStWtResetRel AND #iAutoRunning;
END_REGION

REGION Network 5: STATE Num:0 Reset Released
   RUNG wire#powerrail
      Contact( #sStWtResetRel )
      wire#w1
      I_Contact( #sStWtResetRel_T1 )
      wire#w2
      Coil( #sStWtResetRel )
   END_RUNG
   RUNG wire#powerrail
      I_Contact( #iAutoRunning )
   END_RUNG wire#w1
   RUNG wire#w2
      { S7_GenerateENO := "TRUE" } Move(in := 0, out1 => #StateNo)
   END_RUNG
   // the same network as SCL:
   #sStWtResetRel := (#sStWtResetRel OR NOT #iAutoRunning) AND NOT #sStWtResetRel_T1;
   IF #sStWtResetRel THEN #StateNo := 0; END_IF;
END_REGION

REGION Network 6: Transition for STATE Num:138 Wait for Both Robots Out of Alloy Fixture Center Stand
   RUNG wire#powerrail
      Contact( #s138_WaitBothRbtOutAl )
      I_Contact( #sStWtResetRel )
      Contact( #sSst )
      wire#w1
      Contact( #iRobotOutofZone )
      I_Contact( #iFixTrayPresent )
      Coil( #s138_WaitBothRbtOutAl_T1 )
   END_RUNG
   RUNG wire#w1
      I_Contact( #s138_WaitBothRbtOutAl_T1 )
      Contact( #iRobotOutofZone )
      Contact( #iFixTrayPresent )
      Coil( #s138_WaitBothRbtOutAl_T2 )
   END_RUNG
   // the same network as SCL:
   #_w1 := #s138_WaitBothRbtOutAl AND NOT #sStWtResetRel AND #sSst;
   #s138_WaitBothRbtOutAl_T1 := #_w1 AND #iRobotOutofZone AND NOT #iFixTrayPresent;
   #s138_WaitBothRbtOutAl_T2 := #_w1 AND NOT #s138_WaitBothRbtOutAl_T1 AND #iRobotOutofZone AND #iFixTrayPresent;
END_REGION

REGION Network 7: STATE Num:138 Wait for Both Robots Out of Alloy Fixture Center Stand
   RUNG wire#powerrail
      Contact( #s138_WaitBothRbtOutAl )
      wire#w1
      I_Contact( #sStWtResetRel )
      I_Contact( #s138_WaitBothRbtOutAl_T1 )
      I_Contact( #s138_WaitBothRbtOutAl_T2 )
      wire#w2
      Coil( #s138_WaitBothRbtOutAl )
   END_RUNG
   RUNG wire#powerrail
      Contact( #s149_RbtPickTrayChkEm_T1 )
   END_RUNG wire#w1
   RUNG wire#powerrail
      Contact( #sStWtResetRel_T1 )
   END_RUNG wire#w1
   RUNG wire#w2
      { S7_GenerateENO := "TRUE" } Move(in := 138, out1 => #StateNo)
   END_RUNG
   // the same network as SCL:
   #s138_WaitBothRbtOutAl := (#s138_WaitBothRbtOutAl OR #s149_RbtPickTrayChkEm_T1 OR #sStWtResetRel_T1) AND NOT #sStWtResetRel AND NOT #s138_WaitBothRbtOutAl_T1 AND NOT #s138_WaitBothRbtOutAl_T2;
   IF #s138_WaitBothRbtOutAl THEN #StateNo := 138; END_IF;
END_REGION

REGION Network 8: Transition for STATE Num:139 Fix Empty
   RUNG wire#powerrail
      Contact( #s139_FixEmpty )
      I_Contact( #sStWtResetRel )
      Contact( #sSst )
      Contact( #iFixEmpty )
      Coil( #s139_FixEmpty_T1 )
   END_RUNG
   // the same network as SCL:
   #s139_FixEmpty_T1 := #s139_FixEmpty AND NOT #sStWtResetRel AND #sSst AND #iFixEmpty;
END_REGION

REGION Network 9: STATE Num:139 Fix Empty
   RUNG wire#powerrail
      Contact( #s139_FixEmpty )
      wire#w1
      I_Contact( #sStWtResetRel )
      I_Contact( #s139_FixEmpty_T1 )
      wire#w2
      Coil( #s139_FixEmpty )
   END_RUNG
   RUNG wire#powerrail
      Contact( #s138_WaitBothRbtOutAl_T1 )
   END_RUNG wire#w1
   RUNG wire#w2
      { S7_GenerateENO := "TRUE" } Move(in := 139, out1 => #StateNo)
   END_RUNG
   // the same network as SCL:
   #s139_FixEmpty := (#s139_FixEmpty OR #s138_WaitBothRbtOutAl_T1) AND NOT #sStWtResetRel AND NOT #s139_FixEmpty_T1;
   IF #s139_FixEmpty THEN #StateNo := 139; END_IF;
END_REGION

REGION Network 10: Transition for STATE Num:140 Fix Tray Present_Rec Operation pending
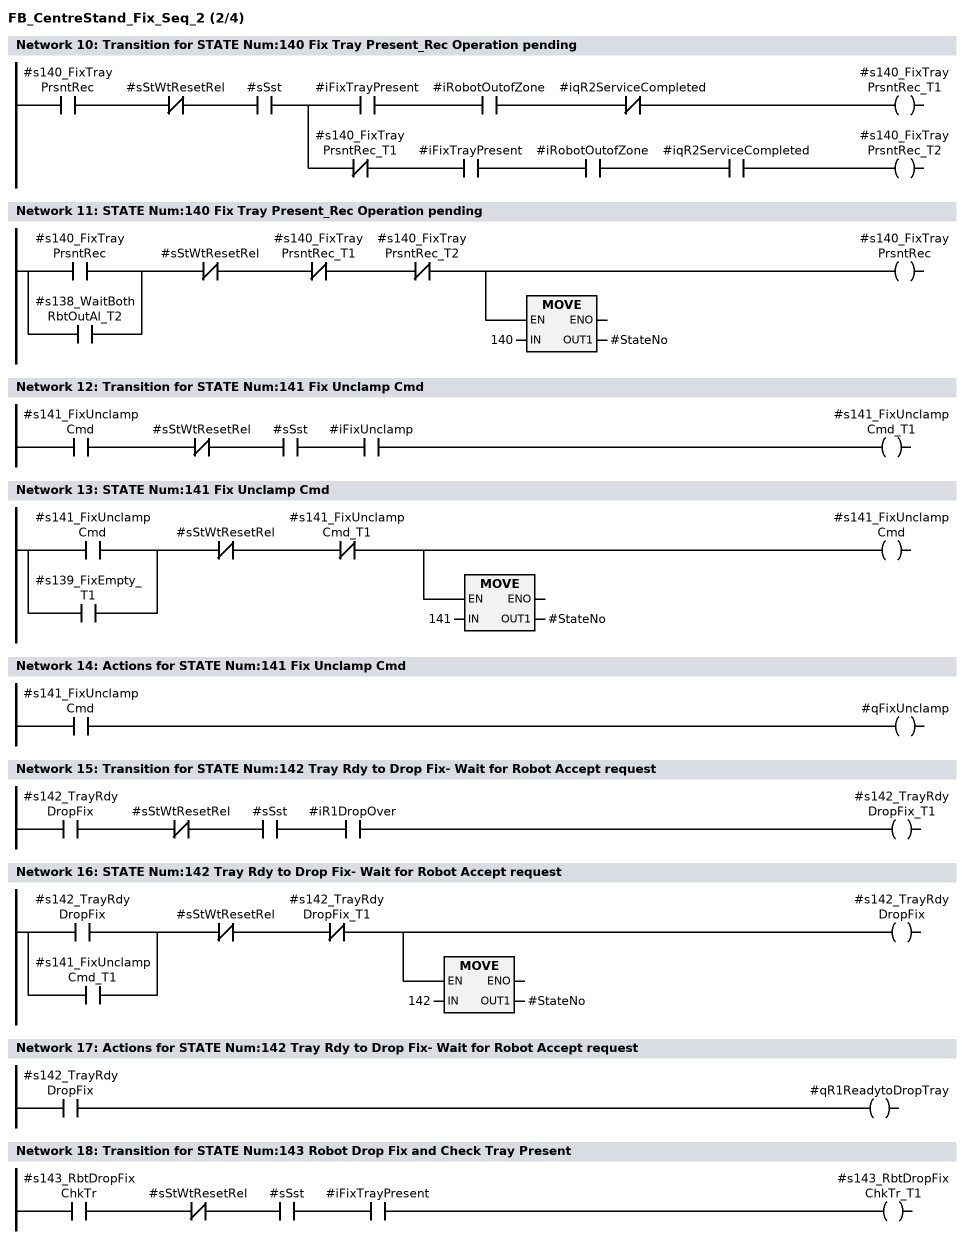
   RUNG wire#powerrail
      Contact( #s140_FixTrayPrsntRec )
      I_Contact( #sStWtResetRel )
      Contact( #sSst )
      wire#w1
      Contact( #iFixTrayPresent )
      Contact( #iRobotOutofZone )
      I_Contact( #iqR2ServiceCompleted )
      Coil( #s140_FixTrayPrsntRec_T1 )
   END_RUNG
   RUNG wire#w1
      I_Contact( #s140_FixTrayPrsntRec_T1 )
      Contact( #iFixTrayPresent )
      Contact( #iRobotOutofZone )
      Contact( #iqR2ServiceCompleted )
      Coil( #s140_FixTrayPrsntRec_T2 )
   END_RUNG
   // the same network as SCL:
   #_w1 := #s140_FixTrayPrsntRec AND NOT #sStWtResetRel AND #sSst;
   #s140_FixTrayPrsntRec_T1 := #_w1 AND #iFixTrayPresent AND #iRobotOutofZone AND NOT #iqR2ServiceCompleted;
   #s140_FixTrayPrsntRec_T2 := #_w1 AND NOT #s140_FixTrayPrsntRec_T1 AND #iFixTrayPresent AND #iRobotOutofZone AND #iqR2ServiceCompleted;
END_REGION

REGION Network 11: STATE Num:140 Fix Tray Present_Rec Operation pending
   RUNG wire#powerrail
      Contact( #s140_FixTrayPrsntRec )
      wire#w1
      I_Contact( #sStWtResetRel )
      I_Contact( #s140_FixTrayPrsntRec_T1 )
      I_Contact( #s140_FixTrayPrsntRec_T2 )
      wire#w2
      Coil( #s140_FixTrayPrsntRec )
   END_RUNG
   RUNG wire#powerrail
      Contact( #s138_WaitBothRbtOutAl_T2 )
   END_RUNG wire#w1
   RUNG wire#w2
      { S7_GenerateENO := "TRUE" } Move(in := 140, out1 => #StateNo)
   END_RUNG
   // the same network as SCL:
   #s140_FixTrayPrsntRec := (#s140_FixTrayPrsntRec OR #s138_WaitBothRbtOutAl_T2) AND NOT #sStWtResetRel AND NOT #s140_FixTrayPrsntRec_T1 AND NOT #s140_FixTrayPrsntRec_T2;
   IF #s140_FixTrayPrsntRec THEN #StateNo := 140; END_IF;
END_REGION

REGION Network 12: Transition for STATE Num:141 Fix Unclamp Cmd
   RUNG wire#powerrail
      Contact( #s141_FixUnclampCmd )
      I_Contact( #sStWtResetRel )
      Contact( #sSst )
      Contact( #iFixUnclamp )
      Coil( #s141_FixUnclampCmd_T1 )
   END_RUNG
   // the same network as SCL:
   #s141_FixUnclampCmd_T1 := #s141_FixUnclampCmd AND NOT #sStWtResetRel AND #sSst AND #iFixUnclamp;
END_REGION

REGION Network 13: STATE Num:141 Fix Unclamp Cmd
   RUNG wire#powerrail
      Contact( #s141_FixUnclampCmd )
      wire#w1
      I_Contact( #sStWtResetRel )
      I_Contact( #s141_FixUnclampCmd_T1 )
      wire#w2
      Coil( #s141_FixUnclampCmd )
   END_RUNG
   RUNG wire#powerrail
      Contact( #s139_FixEmpty_T1 )
   END_RUNG wire#w1
   RUNG wire#w2
      { S7_GenerateENO := "TRUE" } Move(in := 141, out1 => #StateNo)
   END_RUNG
   // the same network as SCL:
   #s141_FixUnclampCmd := (#s141_FixUnclampCmd OR #s139_FixEmpty_T1) AND NOT #sStWtResetRel AND NOT #s141_FixUnclampCmd_T1;
   IF #s141_FixUnclampCmd THEN #StateNo := 141; END_IF;
END_REGION

REGION Network 14: Actions for STATE Num:141 Fix Unclamp Cmd
   RUNG wire#powerrail
      Contact( #s141_FixUnclampCmd )
      Coil( #qFixUnclamp )
   END_RUNG
   // the same network as SCL:
   #qFixUnclamp := #s141_FixUnclampCmd;
END_REGION

REGION Network 15: Transition for STATE Num:142 Tray Rdy to Drop Fix- Wait for Robot Accept request
   RUNG wire#powerrail
      Contact( #s142_TrayRdyDropFix )
      I_Contact( #sStWtResetRel )
      Contact( #sSst )
      Contact( #iR1DropOver )
      Coil( #s142_TrayRdyDropFix_T1 )
   END_RUNG
   // the same network as SCL:
   #s142_TrayRdyDropFix_T1 := #s142_TrayRdyDropFix AND NOT #sStWtResetRel AND #sSst AND #iR1DropOver;
END_REGION

REGION Network 16: STATE Num:142 Tray Rdy to Drop Fix- Wait for Robot Accept request
   RUNG wire#powerrail
      Contact( #s142_TrayRdyDropFix )
      wire#w1
      I_Contact( #sStWtResetRel )
      I_Contact( #s142_TrayRdyDropFix_T1 )
      wire#w2
      Coil( #s142_TrayRdyDropFix )
   END_RUNG
   RUNG wire#powerrail
      Contact( #s141_FixUnclampCmd_T1 )
   END_RUNG wire#w1
   RUNG wire#w2
      { S7_GenerateENO := "TRUE" } Move(in := 142, out1 => #StateNo)
   END_RUNG
   // the same network as SCL:
   #s142_TrayRdyDropFix := (#s142_TrayRdyDropFix OR #s141_FixUnclampCmd_T1) AND NOT #sStWtResetRel AND NOT #s142_TrayRdyDropFix_T1;
   IF #s142_TrayRdyDropFix THEN #StateNo := 142; END_IF;
END_REGION

REGION Network 17: Actions for STATE Num:142 Tray Rdy to Drop Fix- Wait for Robot Accept request
   RUNG wire#powerrail
      Contact( #s142_TrayRdyDropFix )
      Coil( #qR1ReadytoDropTray )
   END_RUNG
   // the same network as SCL:
   #qR1ReadytoDropTray := #s142_TrayRdyDropFix;
END_REGION

REGION Network 18: Transition for STATE Num:143 Robot Drop Fix and Check Tray Present
   RUNG wire#powerrail
      Contact( #s143_RbtDropFixChkTr )
      I_Contact( #sStWtResetRel )
      Contact( #sSst )
      Contact( #iFixTrayPresent )
      Coil( #s143_RbtDropFixChkTr_T1 )
   END_RUNG
   // the same network as SCL:
   #s143_RbtDropFixChkTr_T1 := #s143_RbtDropFixChkTr AND NOT #sStWtResetRel AND #sSst AND #iFixTrayPresent;
END_REGION

REGION Network 19: STATE Num:143 Robot Drop Fix and Check Tray Present
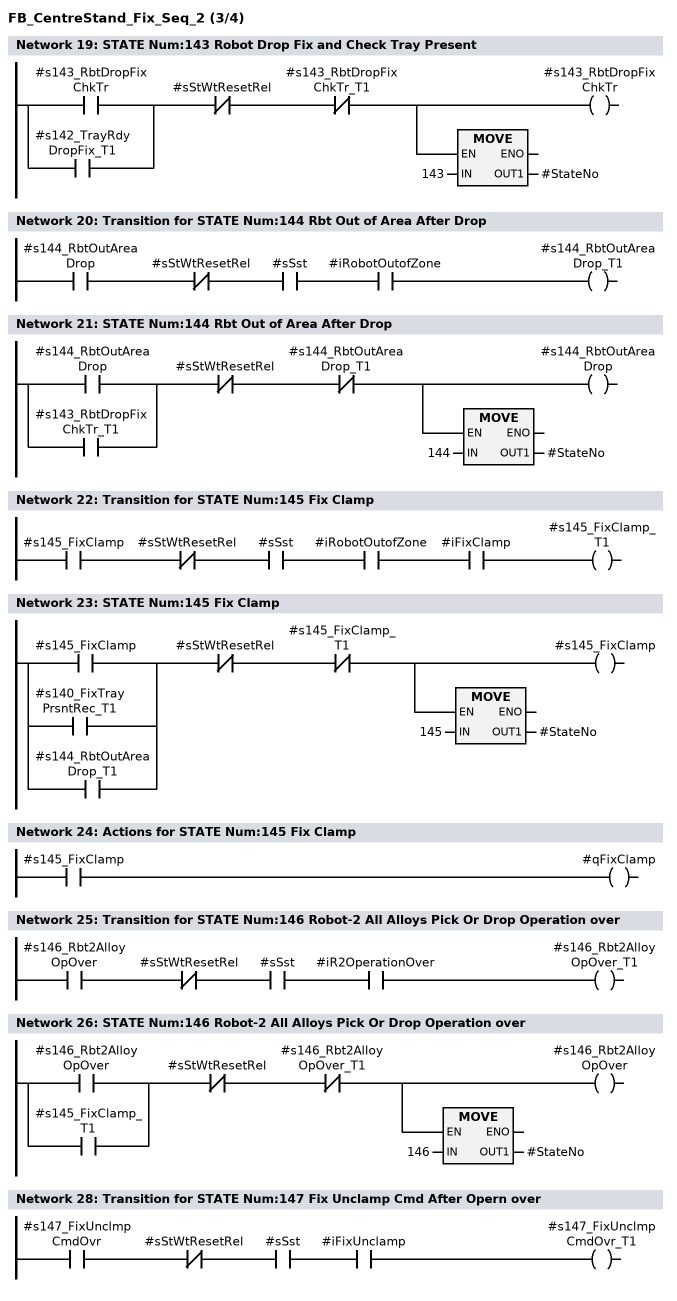
   RUNG wire#powerrail
      Contact( #s143_RbtDropFixChkTr )
      wire#w1
      I_Contact( #sStWtResetRel )
      I_Contact( #s143_RbtDropFixChkTr_T1 )
      wire#w2
      Coil( #s143_RbtDropFixChkTr )
   END_RUNG
   RUNG wire#powerrail
      Contact( #s142_TrayRdyDropFix_T1 )
   END_RUNG wire#w1
   RUNG wire#w2
      { S7_GenerateENO := "TRUE" } Move(in := 143, out1 => #StateNo)
   END_RUNG
   // the same network as SCL:
   #s143_RbtDropFixChkTr := (#s143_RbtDropFixChkTr OR #s142_TrayRdyDropFix_T1) AND NOT #sStWtResetRel AND NOT #s143_RbtDropFixChkTr_T1;
   IF #s143_RbtDropFixChkTr THEN #StateNo := 143; END_IF;
END_REGION

REGION Network 20: Transition for STATE Num:144 Rbt Out of Area After Drop
   RUNG wire#powerrail
      Contact( #s144_RbtOutAreaDrop )
      I_Contact( #sStWtResetRel )
      Contact( #sSst )
      Contact( #iRobotOutofZone )
      Coil( #s144_RbtOutAreaDrop_T1 )
   END_RUNG
   // the same network as SCL:
   #s144_RbtOutAreaDrop_T1 := #s144_RbtOutAreaDrop AND NOT #sStWtResetRel AND #sSst AND #iRobotOutofZone;
END_REGION

REGION Network 21: STATE Num:144 Rbt Out of Area After Drop
   RUNG wire#powerrail
      Contact( #s144_RbtOutAreaDrop )
      wire#w1
      I_Contact( #sStWtResetRel )
      I_Contact( #s144_RbtOutAreaDrop_T1 )
      wire#w2
      Coil( #s144_RbtOutAreaDrop )
   END_RUNG
   RUNG wire#powerrail
      Contact( #s143_RbtDropFixChkTr_T1 )
   END_RUNG wire#w1
   RUNG wire#w2
      { S7_GenerateENO := "TRUE" } Move(in := 144, out1 => #StateNo)
   END_RUNG
   // the same network as SCL:
   #s144_RbtOutAreaDrop := (#s144_RbtOutAreaDrop OR #s143_RbtDropFixChkTr_T1) AND NOT #sStWtResetRel AND NOT #s144_RbtOutAreaDrop_T1;
   IF #s144_RbtOutAreaDrop THEN #StateNo := 144; END_IF;
END_REGION

REGION Network 22: Transition for STATE Num:145 Fix Clamp
   RUNG wire#powerrail
      Contact( #s145_FixClamp )
      I_Contact( #sStWtResetRel )
      Contact( #sSst )
      Contact( #iRobotOutofZone )
      Contact( #iFixClamp )
      Coil( #s145_FixClamp_T1 )
   END_RUNG
   // the same network as SCL:
   #s145_FixClamp_T1 := #s145_FixClamp AND NOT #sStWtResetRel AND #sSst AND #iRobotOutofZone AND #iFixClamp;
END_REGION

REGION Network 23: STATE Num:145 Fix Clamp
   RUNG wire#powerrail
      Contact( #s145_FixClamp )
      wire#w1
      I_Contact( #sStWtResetRel )
      I_Contact( #s145_FixClamp_T1 )
      wire#w2
      Coil( #s145_FixClamp )
   END_RUNG
   RUNG wire#powerrail
      Contact( #s140_FixTrayPrsntRec_T1 )
   END_RUNG wire#w1
   RUNG wire#powerrail
      Contact( #s144_RbtOutAreaDrop_T1 )
   END_RUNG wire#w1
   RUNG wire#w2
      { S7_GenerateENO := "TRUE" } Move(in := 145, out1 => #StateNo)
   END_RUNG
   // the same network as SCL:
   #s145_FixClamp := (#s145_FixClamp OR #s140_FixTrayPrsntRec_T1 OR #s144_RbtOutAreaDrop_T1) AND NOT #sStWtResetRel AND NOT #s145_FixClamp_T1;
   IF #s145_FixClamp THEN #StateNo := 145; END_IF;
END_REGION

REGION Network 24: Actions for STATE Num:145 Fix Clamp
   RUNG wire#powerrail
      Contact( #s145_FixClamp )
      Coil( #qFixClamp )
   END_RUNG
   // the same network as SCL:
   #qFixClamp := #s145_FixClamp;
END_REGION

REGION Network 25: Transition for STATE Num:146 Robot-2 All Alloys Pick Or Drop Operation over
   RUNG wire#powerrail
      Contact( #s146_Rbt2AlloyOpOver )
      I_Contact( #sStWtResetRel )
      Contact( #sSst )
      Contact( #iR2OperationOver )
      Coil( #s146_Rbt2AlloyOpOver_T1 )
   END_RUNG
   // the same network as SCL:
   #s146_Rbt2AlloyOpOver_T1 := #s146_Rbt2AlloyOpOver AND NOT #sStWtResetRel AND #sSst AND #iR2OperationOver;
END_REGION

REGION Network 26: STATE Num:146 Robot-2 All Alloys Pick Or Drop Operation over
   RUNG wire#powerrail
      Contact( #s146_Rbt2AlloyOpOver )
      wire#w1
      I_Contact( #sStWtResetRel )
      I_Contact( #s146_Rbt2AlloyOpOver_T1 )
      wire#w2
      Coil( #s146_Rbt2AlloyOpOver )
   END_RUNG
   RUNG wire#powerrail
      Contact( #s145_FixClamp_T1 )
   END_RUNG wire#w1
   RUNG wire#w2
      { S7_GenerateENO := "TRUE" } Move(in := 146, out1 => #StateNo)
   END_RUNG
   // the same network as SCL:
   #s146_Rbt2AlloyOpOver := (#s146_Rbt2AlloyOpOver OR #s145_FixClamp_T1) AND NOT #sStWtResetRel AND NOT #s146_Rbt2AlloyOpOver_T1;
   IF #s146_Rbt2AlloyOpOver THEN #StateNo := 146; END_IF;
END_REGION

REGION Network 27 (STL): Actions for STATE Num:146 Robot-2 All Alloys Pick Or Drop Operation over
         A     #s146_Rbt2AlloyOpOver;
         =     #qR2OperationStart;
         A     #iR2ServiceActivated;
         S     #iqR2ServiceActive;
         A     #iR2OperationOver;
         A     #iqR2ServiceActive;
         R     #iqR2ServiceActive;
END_REGION

REGION Network 28: Transition for STATE Num:147 Fix Unclamp Cmd After Opern over
   RUNG wire#powerrail
      Contact( #s147_FixUnclmpCmdOvr )
      I_Contact( #sStWtResetRel )
      Contact( #sSst )
      Contact( #iFixUnclamp )
      Coil( #s147_FixUnclmpCmdOvr_T1 )
   END_RUNG
   // the same network as SCL:
   #s147_FixUnclmpCmdOvr_T1 := #s147_FixUnclmpCmdOvr AND NOT #sStWtResetRel AND #sSst AND #iFixUnclamp;
END_REGION

REGION Network 29: STATE Num:147 Fix Unclamp Cmd After Opern over
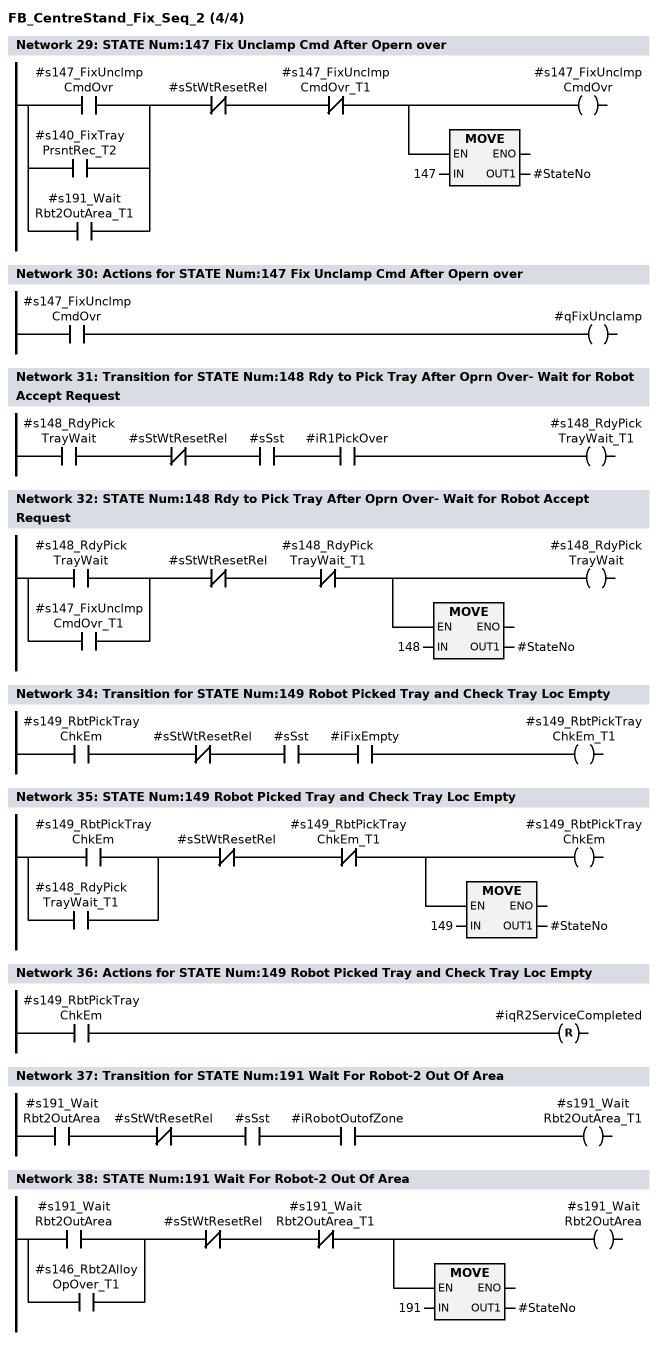
   RUNG wire#powerrail
      Contact( #s147_FixUnclmpCmdOvr )
      wire#w1
      I_Contact( #sStWtResetRel )
      I_Contact( #s147_FixUnclmpCmdOvr_T1 )
      wire#w2
      Coil( #s147_FixUnclmpCmdOvr )
   END_RUNG
   RUNG wire#powerrail
      Contact( #s140_FixTrayPrsntRec_T2 )
   END_RUNG wire#w1
   RUNG wire#powerrail
      Contact( #s191_WaitRbt2OutArea_T1 )
   END_RUNG wire#w1
   RUNG wire#w2
      { S7_GenerateENO := "TRUE" } Move(in := 147, out1 => #StateNo)
   END_RUNG
   // the same network as SCL:
   #s147_FixUnclmpCmdOvr := (#s147_FixUnclmpCmdOvr OR #s140_FixTrayPrsntRec_T2 OR #s191_WaitRbt2OutArea_T1) AND NOT #sStWtResetRel AND NOT #s147_FixUnclmpCmdOvr_T1;
   IF #s147_FixUnclmpCmdOvr THEN #StateNo := 147; END_IF;
END_REGION

REGION Network 30: Actions for STATE Num:147 Fix Unclamp Cmd After Opern over
   RUNG wire#powerrail
      Contact( #s147_FixUnclmpCmdOvr )
      Coil( #qFixUnclamp )
   END_RUNG
   // the same network as SCL:
   #qFixUnclamp := #s147_FixUnclmpCmdOvr;
END_REGION

REGION Network 31: Transition for STATE Num:148 Rdy to Pick Tray After Oprn Over- Wait for Robot Accept Request
   RUNG wire#powerrail
      Contact( #s148_RdyPickTrayWait )
      I_Contact( #sStWtResetRel )
      Contact( #sSst )
      Contact( #iR1PickOver )
      Coil( #s148_RdyPickTrayWait_T1 )
   END_RUNG
   // the same network as SCL:
   #s148_RdyPickTrayWait_T1 := #s148_RdyPickTrayWait AND NOT #sStWtResetRel AND #sSst AND #iR1PickOver;
END_REGION

REGION Network 32: STATE Num:148 Rdy to Pick Tray After Oprn Over- Wait for Robot Accept Request
   RUNG wire#powerrail
      Contact( #s148_RdyPickTrayWait )
      wire#w1
      I_Contact( #sStWtResetRel )
      I_Contact( #s148_RdyPickTrayWait_T1 )
      wire#w2
      Coil( #s148_RdyPickTrayWait )
   END_RUNG
   RUNG wire#powerrail
      Contact( #s147_FixUnclmpCmdOvr_T1 )
   END_RUNG wire#w1
   RUNG wire#w2
      { S7_GenerateENO := "TRUE" } Move(in := 148, out1 => #StateNo)
   END_RUNG
   // the same network as SCL:
   #s148_RdyPickTrayWait := (#s148_RdyPickTrayWait OR #s147_FixUnclmpCmdOvr_T1) AND NOT #sStWtResetRel AND NOT #s148_RdyPickTrayWait_T1;
   IF #s148_RdyPickTrayWait THEN #StateNo := 148; END_IF;
END_REGION

REGION Network 33 (STL): Actions for STATE Num:148 Rdy to Pick Tray After Oprn Over- Wait for Robot Accept Request
         A     #s148_RdyPickTrayWait;
         =     #qR1ReadytoPickTray;
         A     #iR1PickOver;
         R     #iqR2ServiceCompleted;
END_REGION

REGION Network 34: Transition for STATE Num:149 Robot Picked Tray and Check Tray Loc Empty
   RUNG wire#powerrail
      Contact( #s149_RbtPickTrayChkEm )
      I_Contact( #sStWtResetRel )
      Contact( #sSst )
      Contact( #iFixEmpty )
      Coil( #s149_RbtPickTrayChkEm_T1 )
   END_RUNG
   // the same network as SCL:
   #s149_RbtPickTrayChkEm_T1 := #s149_RbtPickTrayChkEm AND NOT #sStWtResetRel AND #sSst AND #iFixEmpty;
END_REGION

REGION Network 35: STATE Num:149 Robot Picked Tray and Check Tray Loc Empty
   RUNG wire#powerrail
      Contact( #s149_RbtPickTrayChkEm )
      wire#w1
      I_Contact( #sStWtResetRel )
      I_Contact( #s149_RbtPickTrayChkEm_T1 )
      wire#w2
      Coil( #s149_RbtPickTrayChkEm )
   END_RUNG
   RUNG wire#powerrail
      Contact( #s148_RdyPickTrayWait_T1 )
   END_RUNG wire#w1
   RUNG wire#w2
      { S7_GenerateENO := "TRUE" } Move(in := 149, out1 => #StateNo)
   END_RUNG
   // the same network as SCL:
   #s149_RbtPickTrayChkEm := (#s149_RbtPickTrayChkEm OR #s148_RdyPickTrayWait_T1) AND NOT #sStWtResetRel AND NOT #s149_RbtPickTrayChkEm_T1;
   IF #s149_RbtPickTrayChkEm THEN #StateNo := 149; END_IF;
END_REGION

REGION Network 36: Actions for STATE Num:149 Robot Picked Tray and Check Tray Loc Empty
   RUNG wire#powerrail
      Contact( #s149_RbtPickTrayChkEm )
      R_Coil( #iqR2ServiceCompleted )
   END_RUNG
   // the same network as SCL:
   IF #s149_RbtPickTrayChkEm THEN #iqR2ServiceCompleted := FALSE; END_IF;
END_REGION

REGION Network 37: Transition for STATE Num:191 Wait For Robot-2 Out Of Area
   RUNG wire#powerrail
      Contact( #s191_WaitRbt2OutArea )
      I_Contact( #sStWtResetRel )
      Contact( #sSst )
      Contact( #iRobotOutofZone )
      Coil( #s191_WaitRbt2OutArea_T1 )
   END_RUNG
   // the same network as SCL:
   #s191_WaitRbt2OutArea_T1 := #s191_WaitRbt2OutArea AND NOT #sStWtResetRel AND #sSst AND #iRobotOutofZone;
END_REGION

REGION Network 38: STATE Num:191 Wait For Robot-2 Out Of Area
   RUNG wire#powerrail
      Contact( #s191_WaitRbt2OutArea )
      wire#w1
      I_Contact( #sStWtResetRel )
      I_Contact( #s191_WaitRbt2OutArea_T1 )
      wire#w2
      Coil( #s191_WaitRbt2OutArea )
   END_RUNG
   RUNG wire#powerrail
      Contact( #s146_Rbt2AlloyOpOver_T1 )
   END_RUNG wire#w1
   RUNG wire#w2
      { S7_GenerateENO := "TRUE" } Move(in := 191, out1 => #StateNo)
   END_RUNG
   // the same network as SCL:
   #s191_WaitRbt2OutArea := (#s191_WaitRbt2OutArea OR #s146_Rbt2AlloyOpOver_T1) AND NOT #sStWtResetRel AND NOT #s191_WaitRbt2OutArea_T1;
   IF #s191_WaitRbt2OutArea THEN #StateNo := 191; END_IF;
END_REGION
END_FUNCTION_BLOCK

FUNCTION_BLOCK "FB_CentreStand_Fix_Seq_3"   // FB1, LAD
{ S7_Optimized_Access := 'TRUE' }
VERSION : 0.1
   VAR_INPUT
      iAutoRunning : Bool;
      iFixClamp : Bool;
      iFixEmpty : Bool;
      iFixTrayPresent : Bool;
      iFixUnclamp : Bool;
      iR1DropOver : Bool;
      iR1PickOver : Bool;
      iR2OperationOver : Bool;
      iR2ServiceActivated : Bool;
      iR2ServiceCompleted : Bool;
      iReset_fault : Bool;
      iRobotOutofZone : Bool;
      iSstMode : Bool;
      iSstPB : Bool;
   END_VAR
   VAR_OUTPUT
      qFixClamp : Bool;
      qFixUnclamp : Bool;
      qR1ReadytoDropTray : Bool;
      qR1ReadytoPickTray : Bool;
      qR2OperationStart : Bool;
   END_VAR
   VAR_IN_OUT
      iqR2ServiceActive : Bool;
      iqR2ServiceCompleted : Bool;
   END_VAR
   VAR
      StateNo : Int;
      s138_WaitBothRbtOutAl : Bool;
      s138_WaitBothRbtOutAl_T1 : Bool;
      s138_WaitBothRbtOutAl_T2 : Bool;
      s139_FixEmpty : Bool;
      s139_FixEmpty_T1 : Bool;
      s140_FixTrayPrsntRec : Bool;
      s140_FixTrayPrsntRec_T1 : Bool;
      s140_FixTrayPrsntRec_T2 : Bool;
      s141_FixUnclampCmd : Bool;
      s141_FixUnclampCmd_T1 : Bool;
      s142_TrayRdyDropFix : Bool;
      s142_TrayRdyDropFix_T1 : Bool;
      s143_RbtDropFixChkTr : Bool;
      s143_RbtDropFixChkTr_T1 : Bool;
      s144_RbtOutAreaDrop : Bool;
      s144_RbtOutAreaDrop_T1 : Bool;
      s145_FixClamp : Bool;
      s145_FixClamp_T1 : Bool;
      s146_Rbt2AlloyOpOver : Bool;
      s146_Rbt2AlloyOpOver_T1 : Bool;
      s147_FixUnclmpCmdOvr : Bool;
      s147_FixUnclmpCmdOvr_T1 : Bool;
      s148_RdyPickTrayWait : Bool;
      s148_RdyPickTrayWait_T1 : Bool;
      s149_RbtPickTrayChkEm : Bool;
      s149_RbtPickTrayChkEm_T1 : Bool;
      s191_WaitRbt2OutArea : Bool;
      s191_WaitRbt2OutArea_T1 : Bool;
      sSst : Bool;
      sSstPulse : Bool;
      sSstRise : Bool;
      sStWtResetRel : Bool;
      sStWtResetRel_T1 : Bool;
   END_VAR
   VAR_TEMP
      tOne : Bool;
   END_VAR
   VAR_TEMP   // added for the SCL form of the ladder/FBD networks
      _w1 : Bool;
   END_VAR
BEGIN

REGION Network 1
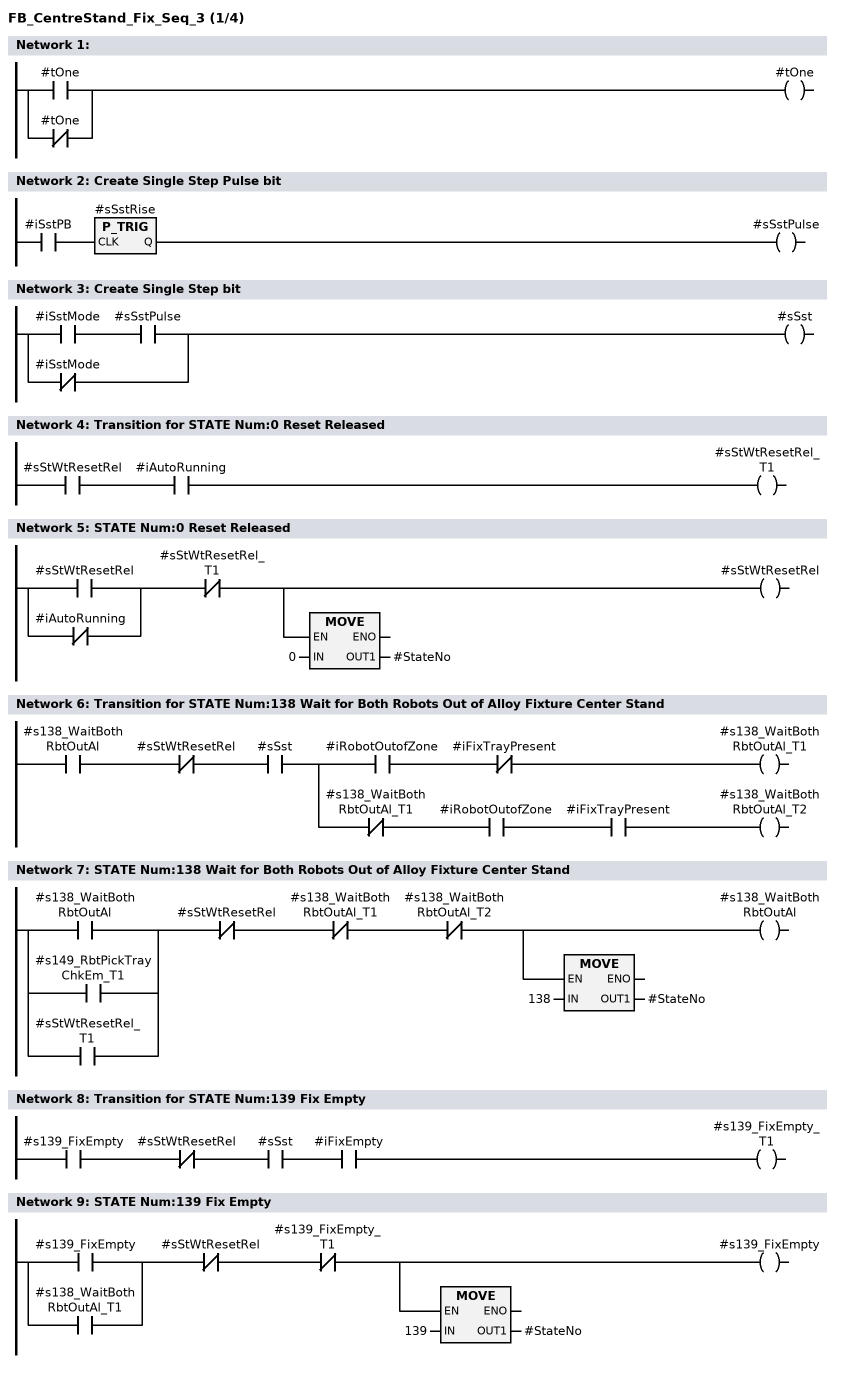
   RUNG wire#powerrail
      Contact( #tOne )
      wire#w1
      Coil( #tOne )
   END_RUNG
   RUNG wire#powerrail
      I_Contact( #tOne )
   END_RUNG wire#w1
   // the same network as SCL:
   #tOne := #tOne OR NOT #tOne;
END_REGION

REGION Network 2: Create Single Step Pulse bit
   RUNG wire#powerrail
      Contact( #iSstPB )
      P_Trig( #sSstRise )
      Coil( #sSstPulse )
   END_RUNG
   // the same network as SCL:
   #_w1 := #iSstPB AND NOT #sSstRise;   // rising edge
   #sSstRise := #iSstPB;
   #sSstPulse := #_w1;
END_REGION

REGION Network 3: Create Single Step bit
   RUNG wire#powerrail
      Contact( #iSstMode )
      Contact( #sSstPulse )
      wire#w1
      Coil( #sSst )
   END_RUNG
   RUNG wire#powerrail
      I_Contact( #iSstMode )
   END_RUNG wire#w1
   // the same network as SCL:
   #sSst := (#iSstMode AND #sSstPulse) OR NOT #iSstMode;
END_REGION

REGION Network 4: Transition for STATE Num:0 Reset Released
   RUNG wire#powerrail
      Contact( #sStWtResetRel )
      Contact( #iAutoRunning )
      Coil( #sStWtResetRel_T1 )
   END_RUNG
   // the same network as SCL:
   #sStWtResetRel_T1 := #sStWtResetRel AND #iAutoRunning;
END_REGION

REGION Network 5: STATE Num:0 Reset Released
   RUNG wire#powerrail
      Contact( #sStWtResetRel )
      wire#w1
      I_Contact( #sStWtResetRel_T1 )
      wire#w2
      Coil( #sStWtResetRel )
   END_RUNG
   RUNG wire#powerrail
      I_Contact( #iAutoRunning )
   END_RUNG wire#w1
   RUNG wire#w2
      { S7_GenerateENO := "TRUE" } Move(in := 0, out1 => #StateNo)
   END_RUNG
   // the same network as SCL:
   #sStWtResetRel := (#sStWtResetRel OR NOT #iAutoRunning) AND NOT #sStWtResetRel_T1;
   IF #sStWtResetRel THEN #StateNo := 0; END_IF;
END_REGION

REGION Network 6: Transition for STATE Num:138 Wait for Both Robots Out of Alloy Fixture Center Stand
   RUNG wire#powerrail
      Contact( #s138_WaitBothRbtOutAl )
      I_Contact( #sStWtResetRel )
      Contact( #sSst )
      wire#w1
      Contact( #iRobotOutofZone )
      I_Contact( #iFixTrayPresent )
      Coil( #s138_WaitBothRbtOutAl_T1 )
   END_RUNG
   RUNG wire#w1
      I_Contact( #s138_WaitBothRbtOutAl_T1 )
      Contact( #iRobotOutofZone )
      Contact( #iFixTrayPresent )
      Coil( #s138_WaitBothRbtOutAl_T2 )
   END_RUNG
   // the same network as SCL:
   #_w1 := #s138_WaitBothRbtOutAl AND NOT #sStWtResetRel AND #sSst;
   #s138_WaitBothRbtOutAl_T1 := #_w1 AND #iRobotOutofZone AND NOT #iFixTrayPresent;
   #s138_WaitBothRbtOutAl_T2 := #_w1 AND NOT #s138_WaitBothRbtOutAl_T1 AND #iRobotOutofZone AND #iFixTrayPresent;
END_REGION

REGION Network 7: STATE Num:138 Wait for Both Robots Out of Alloy Fixture Center Stand
   RUNG wire#powerrail
      Contact( #s138_WaitBothRbtOutAl )
      wire#w1
      I_Contact( #sStWtResetRel )
      I_Contact( #s138_WaitBothRbtOutAl_T1 )
      I_Contact( #s138_WaitBothRbtOutAl_T2 )
      wire#w2
      Coil( #s138_WaitBothRbtOutAl )
   END_RUNG
   RUNG wire#powerrail
      Contact( #s149_RbtPickTrayChkEm_T1 )
   END_RUNG wire#w1
   RUNG wire#powerrail
      Contact( #sStWtResetRel_T1 )
   END_RUNG wire#w1
   RUNG wire#w2
      { S7_GenerateENO := "TRUE" } Move(in := 138, out1 => #StateNo)
   END_RUNG
   // the same network as SCL:
   #s138_WaitBothRbtOutAl := (#s138_WaitBothRbtOutAl OR #s149_RbtPickTrayChkEm_T1 OR #sStWtResetRel_T1) AND NOT #sStWtResetRel AND NOT #s138_WaitBothRbtOutAl_T1 AND NOT #s138_WaitBothRbtOutAl_T2;
   IF #s138_WaitBothRbtOutAl THEN #StateNo := 138; END_IF;
END_REGION

REGION Network 8: Transition for STATE Num:139 Fix Empty
   RUNG wire#powerrail
      Contact( #s139_FixEmpty )
      I_Contact( #sStWtResetRel )
      Contact( #sSst )
      Contact( #iFixEmpty )
      Coil( #s139_FixEmpty_T1 )
   END_RUNG
   // the same network as SCL:
   #s139_FixEmpty_T1 := #s139_FixEmpty AND NOT #sStWtResetRel AND #sSst AND #iFixEmpty;
END_REGION

REGION Network 9: STATE Num:139 Fix Empty
   RUNG wire#powerrail
      Contact( #s139_FixEmpty )
      wire#w1
      I_Contact( #sStWtResetRel )
      I_Contact( #s139_FixEmpty_T1 )
      wire#w2
      Coil( #s139_FixEmpty )
   END_RUNG
   RUNG wire#powerrail
      Contact( #s138_WaitBothRbtOutAl_T1 )
   END_RUNG wire#w1
   RUNG wire#w2
      { S7_GenerateENO := "TRUE" } Move(in := 139, out1 => #StateNo)
   END_RUNG
   // the same network as SCL:
   #s139_FixEmpty := (#s139_FixEmpty OR #s138_WaitBothRbtOutAl_T1) AND NOT #sStWtResetRel AND NOT #s139_FixEmpty_T1;
   IF #s139_FixEmpty THEN #StateNo := 139; END_IF;
END_REGION

REGION Network 10: Transition for STATE Num:140 Fix Tray Present_Rec Operation pending
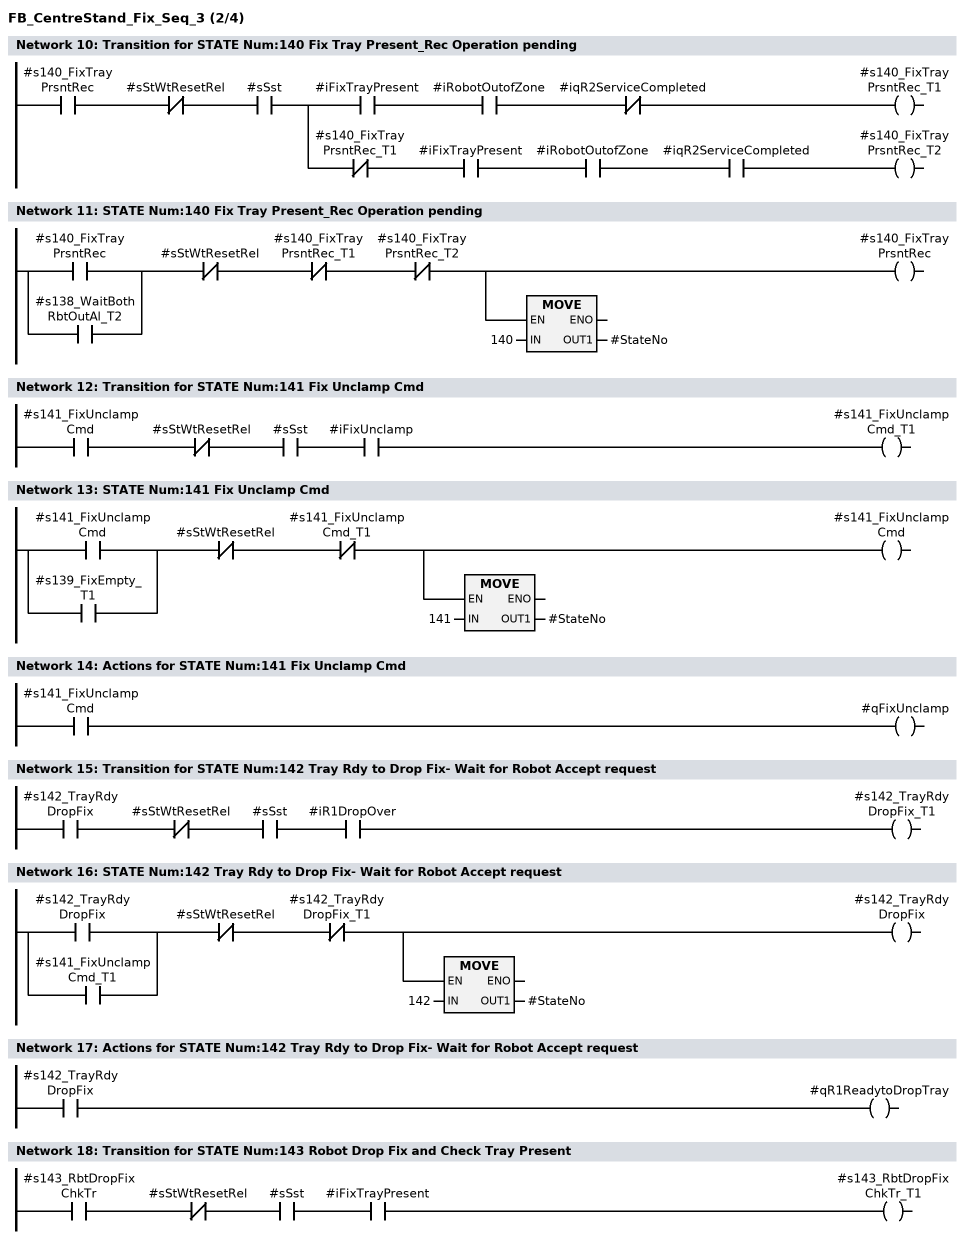
   RUNG wire#powerrail
      Contact( #s140_FixTrayPrsntRec )
      I_Contact( #sStWtResetRel )
      Contact( #sSst )
      wire#w1
      Contact( #iFixTrayPresent )
      Contact( #iRobotOutofZone )
      I_Contact( #iqR2ServiceCompleted )
      Coil( #s140_FixTrayPrsntRec_T1 )
   END_RUNG
   RUNG wire#w1
      I_Contact( #s140_FixTrayPrsntRec_T1 )
      Contact( #iFixTrayPresent )
      Contact( #iRobotOutofZone )
      Contact( #iqR2ServiceCompleted )
      Coil( #s140_FixTrayPrsntRec_T2 )
   END_RUNG
   // the same network as SCL:
   #_w1 := #s140_FixTrayPrsntRec AND NOT #sStWtResetRel AND #sSst;
   #s140_FixTrayPrsntRec_T1 := #_w1 AND #iFixTrayPresent AND #iRobotOutofZone AND NOT #iqR2ServiceCompleted;
   #s140_FixTrayPrsntRec_T2 := #_w1 AND NOT #s140_FixTrayPrsntRec_T1 AND #iFixTrayPresent AND #iRobotOutofZone AND #iqR2ServiceCompleted;
END_REGION

REGION Network 11: STATE Num:140 Fix Tray Present_Rec Operation pending
   RUNG wire#powerrail
      Contact( #s140_FixTrayPrsntRec )
      wire#w1
      I_Contact( #sStWtResetRel )
      I_Contact( #s140_FixTrayPrsntRec_T1 )
      I_Contact( #s140_FixTrayPrsntRec_T2 )
      wire#w2
      Coil( #s140_FixTrayPrsntRec )
   END_RUNG
   RUNG wire#powerrail
      Contact( #s138_WaitBothRbtOutAl_T2 )
   END_RUNG wire#w1
   RUNG wire#w2
      { S7_GenerateENO := "TRUE" } Move(in := 140, out1 => #StateNo)
   END_RUNG
   // the same network as SCL:
   #s140_FixTrayPrsntRec := (#s140_FixTrayPrsntRec OR #s138_WaitBothRbtOutAl_T2) AND NOT #sStWtResetRel AND NOT #s140_FixTrayPrsntRec_T1 AND NOT #s140_FixTrayPrsntRec_T2;
   IF #s140_FixTrayPrsntRec THEN #StateNo := 140; END_IF;
END_REGION

REGION Network 12: Transition for STATE Num:141 Fix Unclamp Cmd
   RUNG wire#powerrail
      Contact( #s141_FixUnclampCmd )
      I_Contact( #sStWtResetRel )
      Contact( #sSst )
      Contact( #iFixUnclamp )
      Coil( #s141_FixUnclampCmd_T1 )
   END_RUNG
   // the same network as SCL:
   #s141_FixUnclampCmd_T1 := #s141_FixUnclampCmd AND NOT #sStWtResetRel AND #sSst AND #iFixUnclamp;
END_REGION

REGION Network 13: STATE Num:141 Fix Unclamp Cmd
   RUNG wire#powerrail
      Contact( #s141_FixUnclampCmd )
      wire#w1
      I_Contact( #sStWtResetRel )
      I_Contact( #s141_FixUnclampCmd_T1 )
      wire#w2
      Coil( #s141_FixUnclampCmd )
   END_RUNG
   RUNG wire#powerrail
      Contact( #s139_FixEmpty_T1 )
   END_RUNG wire#w1
   RUNG wire#w2
      { S7_GenerateENO := "TRUE" } Move(in := 141, out1 => #StateNo)
   END_RUNG
   // the same network as SCL:
   #s141_FixUnclampCmd := (#s141_FixUnclampCmd OR #s139_FixEmpty_T1) AND NOT #sStWtResetRel AND NOT #s141_FixUnclampCmd_T1;
   IF #s141_FixUnclampCmd THEN #StateNo := 141; END_IF;
END_REGION

REGION Network 14: Actions for STATE Num:141 Fix Unclamp Cmd
   RUNG wire#powerrail
      Contact( #s141_FixUnclampCmd )
      Coil( #qFixUnclamp )
   END_RUNG
   // the same network as SCL:
   #qFixUnclamp := #s141_FixUnclampCmd;
END_REGION

REGION Network 15: Transition for STATE Num:142 Tray Rdy to Drop Fix- Wait for Robot Accept request
   RUNG wire#powerrail
      Contact( #s142_TrayRdyDropFix )
      I_Contact( #sStWtResetRel )
      Contact( #sSst )
      Contact( #iR1DropOver )
      Coil( #s142_TrayRdyDropFix_T1 )
   END_RUNG
   // the same network as SCL:
   #s142_TrayRdyDropFix_T1 := #s142_TrayRdyDropFix AND NOT #sStWtResetRel AND #sSst AND #iR1DropOver;
END_REGION

REGION Network 16: STATE Num:142 Tray Rdy to Drop Fix- Wait for Robot Accept request
   RUNG wire#powerrail
      Contact( #s142_TrayRdyDropFix )
      wire#w1
      I_Contact( #sStWtResetRel )
      I_Contact( #s142_TrayRdyDropFix_T1 )
      wire#w2
      Coil( #s142_TrayRdyDropFix )
   END_RUNG
   RUNG wire#powerrail
      Contact( #s141_FixUnclampCmd_T1 )
   END_RUNG wire#w1
   RUNG wire#w2
      { S7_GenerateENO := "TRUE" } Move(in := 142, out1 => #StateNo)
   END_RUNG
   // the same network as SCL:
   #s142_TrayRdyDropFix := (#s142_TrayRdyDropFix OR #s141_FixUnclampCmd_T1) AND NOT #sStWtResetRel AND NOT #s142_TrayRdyDropFix_T1;
   IF #s142_TrayRdyDropFix THEN #StateNo := 142; END_IF;
END_REGION

REGION Network 17: Actions for STATE Num:142 Tray Rdy to Drop Fix- Wait for Robot Accept request
   RUNG wire#powerrail
      Contact( #s142_TrayRdyDropFix )
      Coil( #qR1ReadytoDropTray )
   END_RUNG
   // the same network as SCL:
   #qR1ReadytoDropTray := #s142_TrayRdyDropFix;
END_REGION

REGION Network 18: Transition for STATE Num:143 Robot Drop Fix and Check Tray Present
   RUNG wire#powerrail
      Contact( #s143_RbtDropFixChkTr )
      I_Contact( #sStWtResetRel )
      Contact( #sSst )
      Contact( #iFixTrayPresent )
      Coil( #s143_RbtDropFixChkTr_T1 )
   END_RUNG
   // the same network as SCL:
   #s143_RbtDropFixChkTr_T1 := #s143_RbtDropFixChkTr AND NOT #sStWtResetRel AND #sSst AND #iFixTrayPresent;
END_REGION

REGION Network 19: STATE Num:143 Robot Drop Fix and Check Tray Present
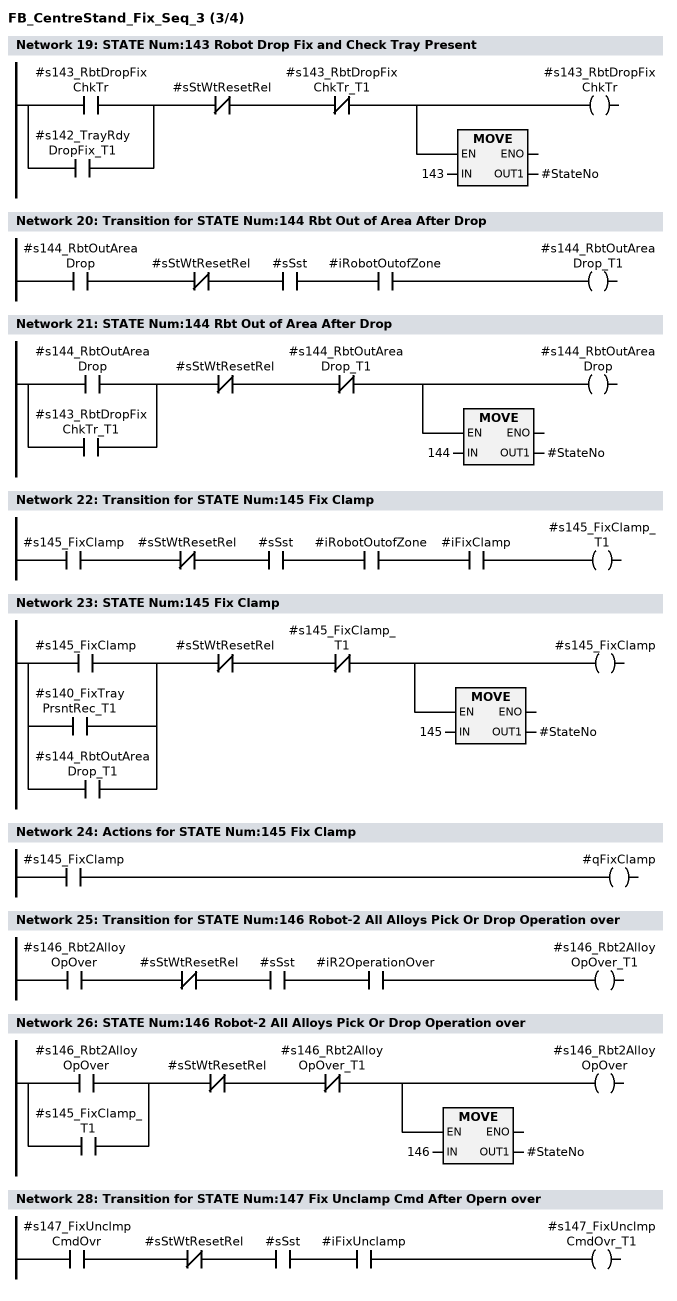
   RUNG wire#powerrail
      Contact( #s143_RbtDropFixChkTr )
      wire#w1
      I_Contact( #sStWtResetRel )
      I_Contact( #s143_RbtDropFixChkTr_T1 )
      wire#w2
      Coil( #s143_RbtDropFixChkTr )
   END_RUNG
   RUNG wire#powerrail
      Contact( #s142_TrayRdyDropFix_T1 )
   END_RUNG wire#w1
   RUNG wire#w2
      { S7_GenerateENO := "TRUE" } Move(in := 143, out1 => #StateNo)
   END_RUNG
   // the same network as SCL:
   #s143_RbtDropFixChkTr := (#s143_RbtDropFixChkTr OR #s142_TrayRdyDropFix_T1) AND NOT #sStWtResetRel AND NOT #s143_RbtDropFixChkTr_T1;
   IF #s143_RbtDropFixChkTr THEN #StateNo := 143; END_IF;
END_REGION

REGION Network 20: Transition for STATE Num:144 Rbt Out of Area After Drop
   RUNG wire#powerrail
      Contact( #s144_RbtOutAreaDrop )
      I_Contact( #sStWtResetRel )
      Contact( #sSst )
      Contact( #iRobotOutofZone )
      Coil( #s144_RbtOutAreaDrop_T1 )
   END_RUNG
   // the same network as SCL:
   #s144_RbtOutAreaDrop_T1 := #s144_RbtOutAreaDrop AND NOT #sStWtResetRel AND #sSst AND #iRobotOutofZone;
END_REGION

REGION Network 21: STATE Num:144 Rbt Out of Area After Drop
   RUNG wire#powerrail
      Contact( #s144_RbtOutAreaDrop )
      wire#w1
      I_Contact( #sStWtResetRel )
      I_Contact( #s144_RbtOutAreaDrop_T1 )
      wire#w2
      Coil( #s144_RbtOutAreaDrop )
   END_RUNG
   RUNG wire#powerrail
      Contact( #s143_RbtDropFixChkTr_T1 )
   END_RUNG wire#w1
   RUNG wire#w2
      { S7_GenerateENO := "TRUE" } Move(in := 144, out1 => #StateNo)
   END_RUNG
   // the same network as SCL:
   #s144_RbtOutAreaDrop := (#s144_RbtOutAreaDrop OR #s143_RbtDropFixChkTr_T1) AND NOT #sStWtResetRel AND NOT #s144_RbtOutAreaDrop_T1;
   IF #s144_RbtOutAreaDrop THEN #StateNo := 144; END_IF;
END_REGION

REGION Network 22: Transition for STATE Num:145 Fix Clamp
   RUNG wire#powerrail
      Contact( #s145_FixClamp )
      I_Contact( #sStWtResetRel )
      Contact( #sSst )
      Contact( #iRobotOutofZone )
      Contact( #iFixClamp )
      Coil( #s145_FixClamp_T1 )
   END_RUNG
   // the same network as SCL:
   #s145_FixClamp_T1 := #s145_FixClamp AND NOT #sStWtResetRel AND #sSst AND #iRobotOutofZone AND #iFixClamp;
END_REGION

REGION Network 23: STATE Num:145 Fix Clamp
   RUNG wire#powerrail
      Contact( #s145_FixClamp )
      wire#w1
      I_Contact( #sStWtResetRel )
      I_Contact( #s145_FixClamp_T1 )
      wire#w2
      Coil( #s145_FixClamp )
   END_RUNG
   RUNG wire#powerrail
      Contact( #s140_FixTrayPrsntRec_T1 )
   END_RUNG wire#w1
   RUNG wire#powerrail
      Contact( #s144_RbtOutAreaDrop_T1 )
   END_RUNG wire#w1
   RUNG wire#w2
      { S7_GenerateENO := "TRUE" } Move(in := 145, out1 => #StateNo)
   END_RUNG
   // the same network as SCL:
   #s145_FixClamp := (#s145_FixClamp OR #s140_FixTrayPrsntRec_T1 OR #s144_RbtOutAreaDrop_T1) AND NOT #sStWtResetRel AND NOT #s145_FixClamp_T1;
   IF #s145_FixClamp THEN #StateNo := 145; END_IF;
END_REGION

REGION Network 24: Actions for STATE Num:145 Fix Clamp
   RUNG wire#powerrail
      Contact( #s145_FixClamp )
      Coil( #qFixClamp )
   END_RUNG
   // the same network as SCL:
   #qFixClamp := #s145_FixClamp;
END_REGION

REGION Network 25: Transition for STATE Num:146 Robot-2 All Alloys Pick Or Drop Operation over
   RUNG wire#powerrail
      Contact( #s146_Rbt2AlloyOpOver )
      I_Contact( #sStWtResetRel )
      Contact( #sSst )
      Contact( #iR2OperationOver )
      Coil( #s146_Rbt2AlloyOpOver_T1 )
   END_RUNG
   // the same network as SCL:
   #s146_Rbt2AlloyOpOver_T1 := #s146_Rbt2AlloyOpOver AND NOT #sStWtResetRel AND #sSst AND #iR2OperationOver;
END_REGION

REGION Network 26: STATE Num:146 Robot-2 All Alloys Pick Or Drop Operation over
   RUNG wire#powerrail
      Contact( #s146_Rbt2AlloyOpOver )
      wire#w1
      I_Contact( #sStWtResetRel )
      I_Contact( #s146_Rbt2AlloyOpOver_T1 )
      wire#w2
      Coil( #s146_Rbt2AlloyOpOver )
   END_RUNG
   RUNG wire#powerrail
      Contact( #s145_FixClamp_T1 )
   END_RUNG wire#w1
   RUNG wire#w2
      { S7_GenerateENO := "TRUE" } Move(in := 146, out1 => #StateNo)
   END_RUNG
   // the same network as SCL:
   #s146_Rbt2AlloyOpOver := (#s146_Rbt2AlloyOpOver OR #s145_FixClamp_T1) AND NOT #sStWtResetRel AND NOT #s146_Rbt2AlloyOpOver_T1;
   IF #s146_Rbt2AlloyOpOver THEN #StateNo := 146; END_IF;
END_REGION

REGION Network 27 (STL): Actions for STATE Num:146 Robot-2 All Alloys Pick Or Drop Operation over
         A     #s146_Rbt2AlloyOpOver;
         =     #qR2OperationStart;
         A     #iR2ServiceActivated;
         S     #iqR2ServiceActive;
         A     #iR2OperationOver;
         A     #iqR2ServiceActive;
         R     #iqR2ServiceActive;
END_REGION

REGION Network 28: Transition for STATE Num:147 Fix Unclamp Cmd After Opern over
   RUNG wire#powerrail
      Contact( #s147_FixUnclmpCmdOvr )
      I_Contact( #sStWtResetRel )
      Contact( #sSst )
      Contact( #iFixUnclamp )
      Coil( #s147_FixUnclmpCmdOvr_T1 )
   END_RUNG
   // the same network as SCL:
   #s147_FixUnclmpCmdOvr_T1 := #s147_FixUnclmpCmdOvr AND NOT #sStWtResetRel AND #sSst AND #iFixUnclamp;
END_REGION

REGION Network 29: STATE Num:147 Fix Unclamp Cmd After Opern over
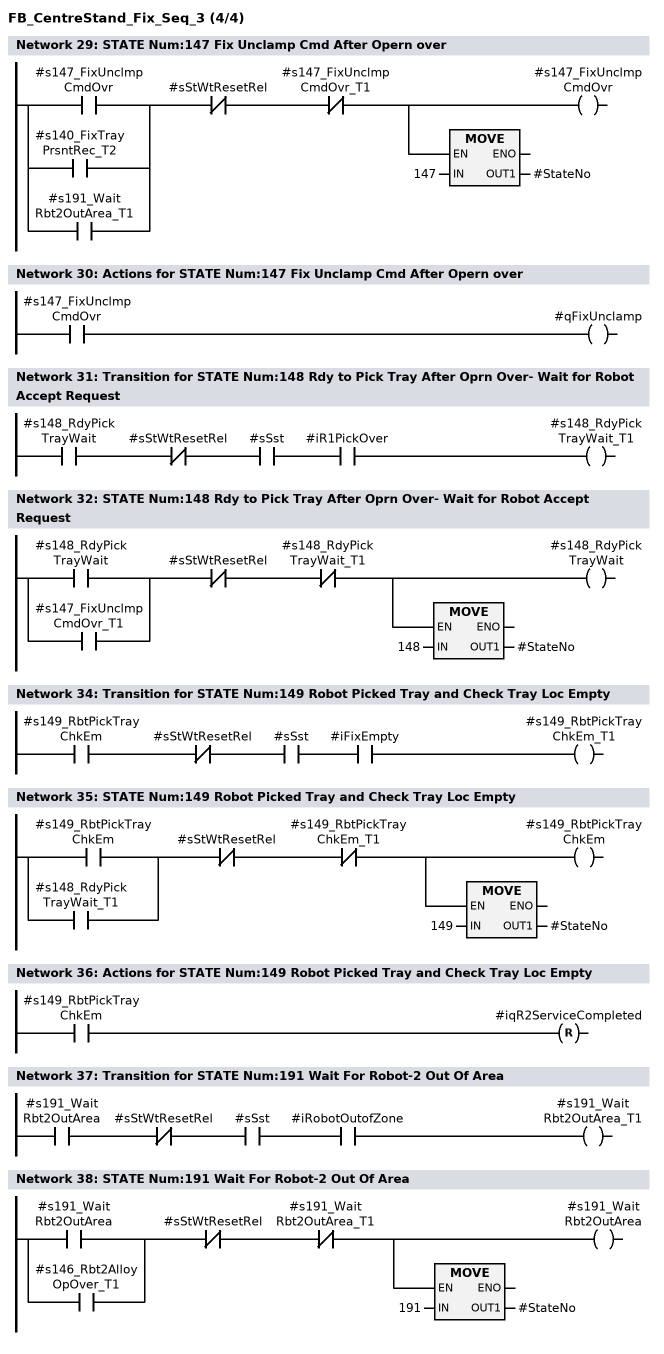
   RUNG wire#powerrail
      Contact( #s147_FixUnclmpCmdOvr )
      wire#w1
      I_Contact( #sStWtResetRel )
      I_Contact( #s147_FixUnclmpCmdOvr_T1 )
      wire#w2
      Coil( #s147_FixUnclmpCmdOvr )
   END_RUNG
   RUNG wire#powerrail
      Contact( #s140_FixTrayPrsntRec_T2 )
   END_RUNG wire#w1
   RUNG wire#powerrail
      Contact( #s191_WaitRbt2OutArea_T1 )
   END_RUNG wire#w1
   RUNG wire#w2
      { S7_GenerateENO := "TRUE" } Move(in := 147, out1 => #StateNo)
   END_RUNG
   // the same network as SCL:
   #s147_FixUnclmpCmdOvr := (#s147_FixUnclmpCmdOvr OR #s140_FixTrayPrsntRec_T2 OR #s191_WaitRbt2OutArea_T1) AND NOT #sStWtResetRel AND NOT #s147_FixUnclmpCmdOvr_T1;
   IF #s147_FixUnclmpCmdOvr THEN #StateNo := 147; END_IF;
END_REGION

REGION Network 30: Actions for STATE Num:147 Fix Unclamp Cmd After Opern over
   RUNG wire#powerrail
      Contact( #s147_FixUnclmpCmdOvr )
      Coil( #qFixUnclamp )
   END_RUNG
   // the same network as SCL:
   #qFixUnclamp := #s147_FixUnclmpCmdOvr;
END_REGION

REGION Network 31: Transition for STATE Num:148 Rdy to Pick Tray After Oprn Over- Wait for Robot Accept Request
   RUNG wire#powerrail
      Contact( #s148_RdyPickTrayWait )
      I_Contact( #sStWtResetRel )
      Contact( #sSst )
      Contact( #iR1PickOver )
      Coil( #s148_RdyPickTrayWait_T1 )
   END_RUNG
   // the same network as SCL:
   #s148_RdyPickTrayWait_T1 := #s148_RdyPickTrayWait AND NOT #sStWtResetRel AND #sSst AND #iR1PickOver;
END_REGION

REGION Network 32: STATE Num:148 Rdy to Pick Tray After Oprn Over- Wait for Robot Accept Request
   RUNG wire#powerrail
      Contact( #s148_RdyPickTrayWait )
      wire#w1
      I_Contact( #sStWtResetRel )
      I_Contact( #s148_RdyPickTrayWait_T1 )
      wire#w2
      Coil( #s148_RdyPickTrayWait )
   END_RUNG
   RUNG wire#powerrail
      Contact( #s147_FixUnclmpCmdOvr_T1 )
   END_RUNG wire#w1
   RUNG wire#w2
      { S7_GenerateENO := "TRUE" } Move(in := 148, out1 => #StateNo)
   END_RUNG
   // the same network as SCL:
   #s148_RdyPickTrayWait := (#s148_RdyPickTrayWait OR #s147_FixUnclmpCmdOvr_T1) AND NOT #sStWtResetRel AND NOT #s148_RdyPickTrayWait_T1;
   IF #s148_RdyPickTrayWait THEN #StateNo := 148; END_IF;
END_REGION

REGION Network 33 (STL): Actions for STATE Num:148 Rdy to Pick Tray After Oprn Over- Wait for Robot Accept Request
         A     #s148_RdyPickTrayWait;
         =     #qR1ReadytoPickTray;
         A     #iR1PickOver;
         R     #iqR2ServiceCompleted;
END_REGION

REGION Network 34: Transition for STATE Num:149 Robot Picked Tray and Check Tray Loc Empty
   RUNG wire#powerrail
      Contact( #s149_RbtPickTrayChkEm )
      I_Contact( #sStWtResetRel )
      Contact( #sSst )
      Contact( #iFixEmpty )
      Coil( #s149_RbtPickTrayChkEm_T1 )
   END_RUNG
   // the same network as SCL:
   #s149_RbtPickTrayChkEm_T1 := #s149_RbtPickTrayChkEm AND NOT #sStWtResetRel AND #sSst AND #iFixEmpty;
END_REGION

REGION Network 35: STATE Num:149 Robot Picked Tray and Check Tray Loc Empty
   RUNG wire#powerrail
      Contact( #s149_RbtPickTrayChkEm )
      wire#w1
      I_Contact( #sStWtResetRel )
      I_Contact( #s149_RbtPickTrayChkEm_T1 )
      wire#w2
      Coil( #s149_RbtPickTrayChkEm )
   END_RUNG
   RUNG wire#powerrail
      Contact( #s148_RdyPickTrayWait_T1 )
   END_RUNG wire#w1
   RUNG wire#w2
      { S7_GenerateENO := "TRUE" } Move(in := 149, out1 => #StateNo)
   END_RUNG
   // the same network as SCL:
   #s149_RbtPickTrayChkEm := (#s149_RbtPickTrayChkEm OR #s148_RdyPickTrayWait_T1) AND NOT #sStWtResetRel AND NOT #s149_RbtPickTrayChkEm_T1;
   IF #s149_RbtPickTrayChkEm THEN #StateNo := 149; END_IF;
END_REGION

REGION Network 36: Actions for STATE Num:149 Robot Picked Tray and Check Tray Loc Empty
   RUNG wire#powerrail
      Contact( #s149_RbtPickTrayChkEm )
      R_Coil( #iqR2ServiceCompleted )
   END_RUNG
   // the same network as SCL:
   IF #s149_RbtPickTrayChkEm THEN #iqR2ServiceCompleted := FALSE; END_IF;
END_REGION

REGION Network 37: Transition for STATE Num:191 Wait For Robot-2 Out Of Area
   RUNG wire#powerrail
      Contact( #s191_WaitRbt2OutArea )
      I_Contact( #sStWtResetRel )
      Contact( #sSst )
      Contact( #iRobotOutofZone )
      Coil( #s191_WaitRbt2OutArea_T1 )
   END_RUNG
   // the same network as SCL:
   #s191_WaitRbt2OutArea_T1 := #s191_WaitRbt2OutArea AND NOT #sStWtResetRel AND #sSst AND #iRobotOutofZone;
END_REGION

REGION Network 38: STATE Num:191 Wait For Robot-2 Out Of Area
   RUNG wire#powerrail
      Contact( #s191_WaitRbt2OutArea )
      wire#w1
      I_Contact( #sStWtResetRel )
      I_Contact( #s191_WaitRbt2OutArea_T1 )
      wire#w2
      Coil( #s191_WaitRbt2OutArea )
   END_RUNG
   RUNG wire#powerrail
      Contact( #s146_Rbt2AlloyOpOver_T1 )
   END_RUNG wire#w1
   RUNG wire#w2
      { S7_GenerateENO := "TRUE" } Move(in := 191, out1 => #StateNo)
   END_RUNG
   // the same network as SCL:
   #s191_WaitRbt2OutArea := (#s191_WaitRbt2OutArea OR #s146_Rbt2AlloyOpOver_T1) AND NOT #sStWtResetRel AND NOT #s191_WaitRbt2OutArea_T1;
   IF #s191_WaitRbt2OutArea THEN #StateNo := 191; END_IF;
END_REGION
END_FUNCTION_BLOCK

FUNCTION_BLOCK "FB_CentreStand_Fix_Seq_4"   // FB1, LAD
{ S7_Optimized_Access := 'TRUE' }
VERSION : 0.1
   VAR_INPUT
      iAutoRunning : Bool;
      iFixClamp : Bool;
      iFixEmpty : Bool;
      iFixTrayPresent : Bool;
      iFixUnclamp : Bool;
      iR1DropOver : Bool;
      iR1PickOver : Bool;
      iR2OperationOver : Bool;
      iR2ServiceActivated : Bool;
      iR2ServiceCompleted : Bool;
      iReset_fault : Bool;
      iRobotOutofZone : Bool;
      iSstMode : Bool;
      iSstPB : Bool;
   END_VAR
   VAR_OUTPUT
      qFixClamp : Bool;
      qFixUnclamp : Bool;
      qR1ReadytoDropTray : Bool;
      qR1ReadytoPickTray : Bool;
      qR2OperationStart : Bool;
   END_VAR
   VAR_IN_OUT
      iqR2ServiceActive : Bool;
      iqR2ServiceCompleted : Bool;
   END_VAR
   VAR
      StateNo : Int;
      s138_WaitBothRbtOutAl : Bool;
      s138_WaitBothRbtOutAl_T1 : Bool;
      s138_WaitBothRbtOutAl_T2 : Bool;
      s139_FixEmpty : Bool;
      s139_FixEmpty_T1 : Bool;
      s140_FixTrayPrsntRec : Bool;
      s140_FixTrayPrsntRec_T1 : Bool;
      s140_FixTrayPrsntRec_T2 : Bool;
      s141_FixUnclampCmd : Bool;
      s141_FixUnclampCmd_T1 : Bool;
      s142_TrayRdyDropFix : Bool;
      s142_TrayRdyDropFix_T1 : Bool;
      s143_RbtDropFixChkTr : Bool;
      s143_RbtDropFixChkTr_T1 : Bool;
      s144_RbtOutAreaDrop : Bool;
      s144_RbtOutAreaDrop_T1 : Bool;
      s145_FixClamp : Bool;
      s145_FixClamp_T1 : Bool;
      s146_Rbt2AlloyOpOver : Bool;
      s146_Rbt2AlloyOpOver_T1 : Bool;
      s147_FixUnclmpCmdOvr : Bool;
      s147_FixUnclmpCmdOvr_T1 : Bool;
      s148_RdyPickTrayWait : Bool;
      s148_RdyPickTrayWait_T1 : Bool;
      s149_RbtPickTrayChkEm : Bool;
      s149_RbtPickTrayChkEm_T1 : Bool;
      s191_WaitRbt2OutArea : Bool;
      s191_WaitRbt2OutArea_T1 : Bool;
      sSst : Bool;
      sSstPulse : Bool;
      sSstRise : Bool;
      sStWtResetRel : Bool;
      sStWtResetRel_T1 : Bool;
   END_VAR
   VAR_TEMP
      tOne : Bool;
   END_VAR
   VAR_TEMP   // added for the SCL form of the ladder/FBD networks
      _w1 : Bool;
   END_VAR
BEGIN

REGION Network 1
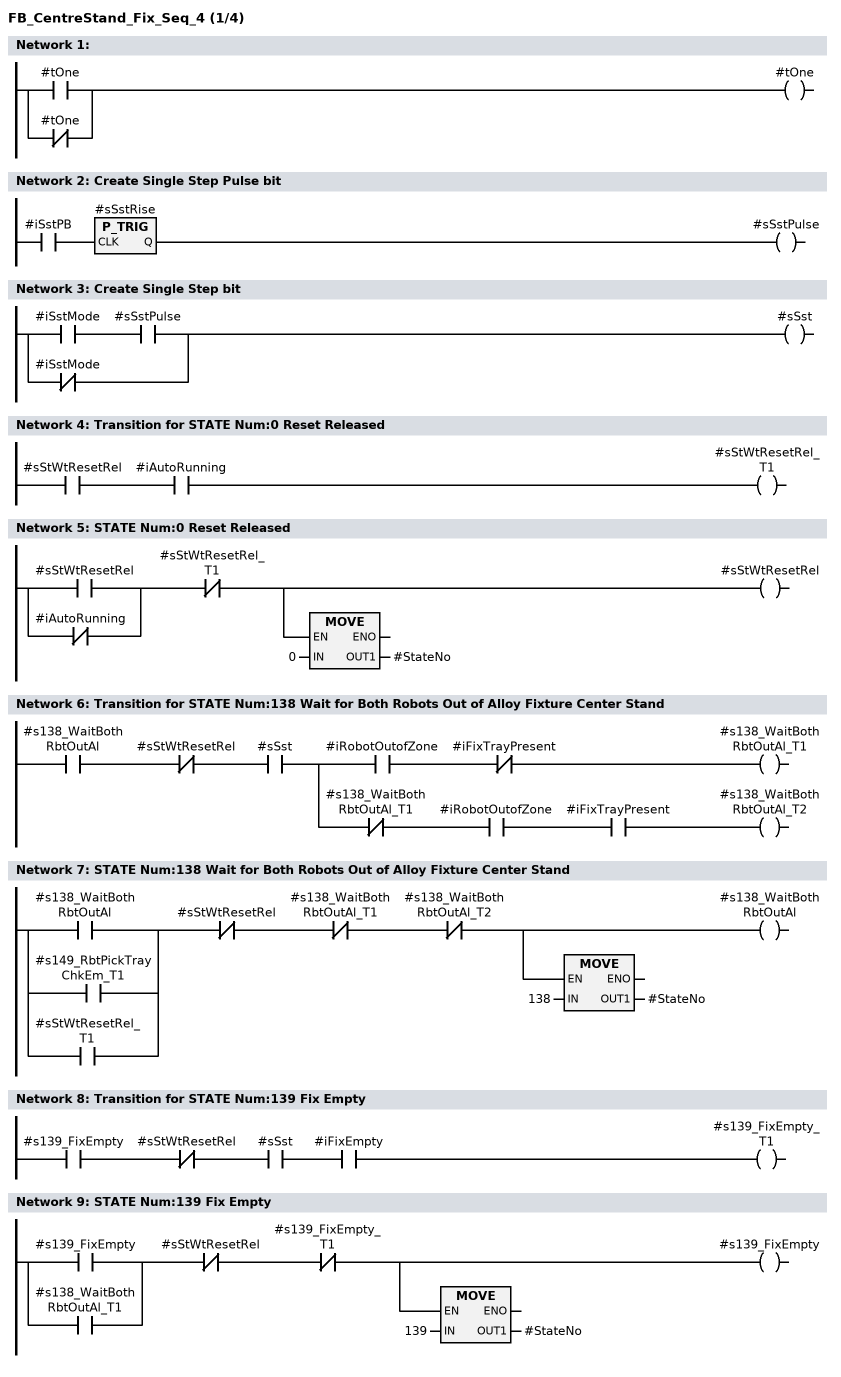
   RUNG wire#powerrail
      Contact( #tOne )
      wire#w1
      Coil( #tOne )
   END_RUNG
   RUNG wire#powerrail
      I_Contact( #tOne )
   END_RUNG wire#w1
   // the same network as SCL:
   #tOne := #tOne OR NOT #tOne;
END_REGION

REGION Network 2: Create Single Step Pulse bit
   RUNG wire#powerrail
      Contact( #iSstPB )
      P_Trig( #sSstRise )
      Coil( #sSstPulse )
   END_RUNG
   // the same network as SCL:
   #_w1 := #iSstPB AND NOT #sSstRise;   // rising edge
   #sSstRise := #iSstPB;
   #sSstPulse := #_w1;
END_REGION

REGION Network 3: Create Single Step bit
   RUNG wire#powerrail
      Contact( #iSstMode )
      Contact( #sSstPulse )
      wire#w1
      Coil( #sSst )
   END_RUNG
   RUNG wire#powerrail
      I_Contact( #iSstMode )
   END_RUNG wire#w1
   // the same network as SCL:
   #sSst := (#iSstMode AND #sSstPulse) OR NOT #iSstMode;
END_REGION

REGION Network 4: Transition for STATE Num:0 Reset Released
   RUNG wire#powerrail
      Contact( #sStWtResetRel )
      Contact( #iAutoRunning )
      Coil( #sStWtResetRel_T1 )
   END_RUNG
   // the same network as SCL:
   #sStWtResetRel_T1 := #sStWtResetRel AND #iAutoRunning;
END_REGION

REGION Network 5: STATE Num:0 Reset Released
   RUNG wire#powerrail
      Contact( #sStWtResetRel )
      wire#w1
      I_Contact( #sStWtResetRel_T1 )
      wire#w2
      Coil( #sStWtResetRel )
   END_RUNG
   RUNG wire#powerrail
      I_Contact( #iAutoRunning )
   END_RUNG wire#w1
   RUNG wire#w2
      { S7_GenerateENO := "TRUE" } Move(in := 0, out1 => #StateNo)
   END_RUNG
   // the same network as SCL:
   #sStWtResetRel := (#sStWtResetRel OR NOT #iAutoRunning) AND NOT #sStWtResetRel_T1;
   IF #sStWtResetRel THEN #StateNo := 0; END_IF;
END_REGION

REGION Network 6: Transition for STATE Num:138 Wait for Both Robots Out of Alloy Fixture Center Stand
   RUNG wire#powerrail
      Contact( #s138_WaitBothRbtOutAl )
      I_Contact( #sStWtResetRel )
      Contact( #sSst )
      wire#w1
      Contact( #iRobotOutofZone )
      I_Contact( #iFixTrayPresent )
      Coil( #s138_WaitBothRbtOutAl_T1 )
   END_RUNG
   RUNG wire#w1
      I_Contact( #s138_WaitBothRbtOutAl_T1 )
      Contact( #iRobotOutofZone )
      Contact( #iFixTrayPresent )
      Coil( #s138_WaitBothRbtOutAl_T2 )
   END_RUNG
   // the same network as SCL:
   #_w1 := #s138_WaitBothRbtOutAl AND NOT #sStWtResetRel AND #sSst;
   #s138_WaitBothRbtOutAl_T1 := #_w1 AND #iRobotOutofZone AND NOT #iFixTrayPresent;
   #s138_WaitBothRbtOutAl_T2 := #_w1 AND NOT #s138_WaitBothRbtOutAl_T1 AND #iRobotOutofZone AND #iFixTrayPresent;
END_REGION

REGION Network 7: STATE Num:138 Wait for Both Robots Out of Alloy Fixture Center Stand
   RUNG wire#powerrail
      Contact( #s138_WaitBothRbtOutAl )
      wire#w1
      I_Contact( #sStWtResetRel )
      I_Contact( #s138_WaitBothRbtOutAl_T1 )
      I_Contact( #s138_WaitBothRbtOutAl_T2 )
      wire#w2
      Coil( #s138_WaitBothRbtOutAl )
   END_RUNG
   RUNG wire#powerrail
      Contact( #s149_RbtPickTrayChkEm_T1 )
   END_RUNG wire#w1
   RUNG wire#powerrail
      Contact( #sStWtResetRel_T1 )
   END_RUNG wire#w1
   RUNG wire#w2
      { S7_GenerateENO := "TRUE" } Move(in := 138, out1 => #StateNo)
   END_RUNG
   // the same network as SCL:
   #s138_WaitBothRbtOutAl := (#s138_WaitBothRbtOutAl OR #s149_RbtPickTrayChkEm_T1 OR #sStWtResetRel_T1) AND NOT #sStWtResetRel AND NOT #s138_WaitBothRbtOutAl_T1 AND NOT #s138_WaitBothRbtOutAl_T2;
   IF #s138_WaitBothRbtOutAl THEN #StateNo := 138; END_IF;
END_REGION

REGION Network 8: Transition for STATE Num:139 Fix Empty
   RUNG wire#powerrail
      Contact( #s139_FixEmpty )
      I_Contact( #sStWtResetRel )
      Contact( #sSst )
      Contact( #iFixEmpty )
      Coil( #s139_FixEmpty_T1 )
   END_RUNG
   // the same network as SCL:
   #s139_FixEmpty_T1 := #s139_FixEmpty AND NOT #sStWtResetRel AND #sSst AND #iFixEmpty;
END_REGION

REGION Network 9: STATE Num:139 Fix Empty
   RUNG wire#powerrail
      Contact( #s139_FixEmpty )
      wire#w1
      I_Contact( #sStWtResetRel )
      I_Contact( #s139_FixEmpty_T1 )
      wire#w2
      Coil( #s139_FixEmpty )
   END_RUNG
   RUNG wire#powerrail
      Contact( #s138_WaitBothRbtOutAl_T1 )
   END_RUNG wire#w1
   RUNG wire#w2
      { S7_GenerateENO := "TRUE" } Move(in := 139, out1 => #StateNo)
   END_RUNG
   // the same network as SCL:
   #s139_FixEmpty := (#s139_FixEmpty OR #s138_WaitBothRbtOutAl_T1) AND NOT #sStWtResetRel AND NOT #s139_FixEmpty_T1;
   IF #s139_FixEmpty THEN #StateNo := 139; END_IF;
END_REGION

REGION Network 10: Transition for STATE Num:140 Fix Tray Present_Rec Operation pending
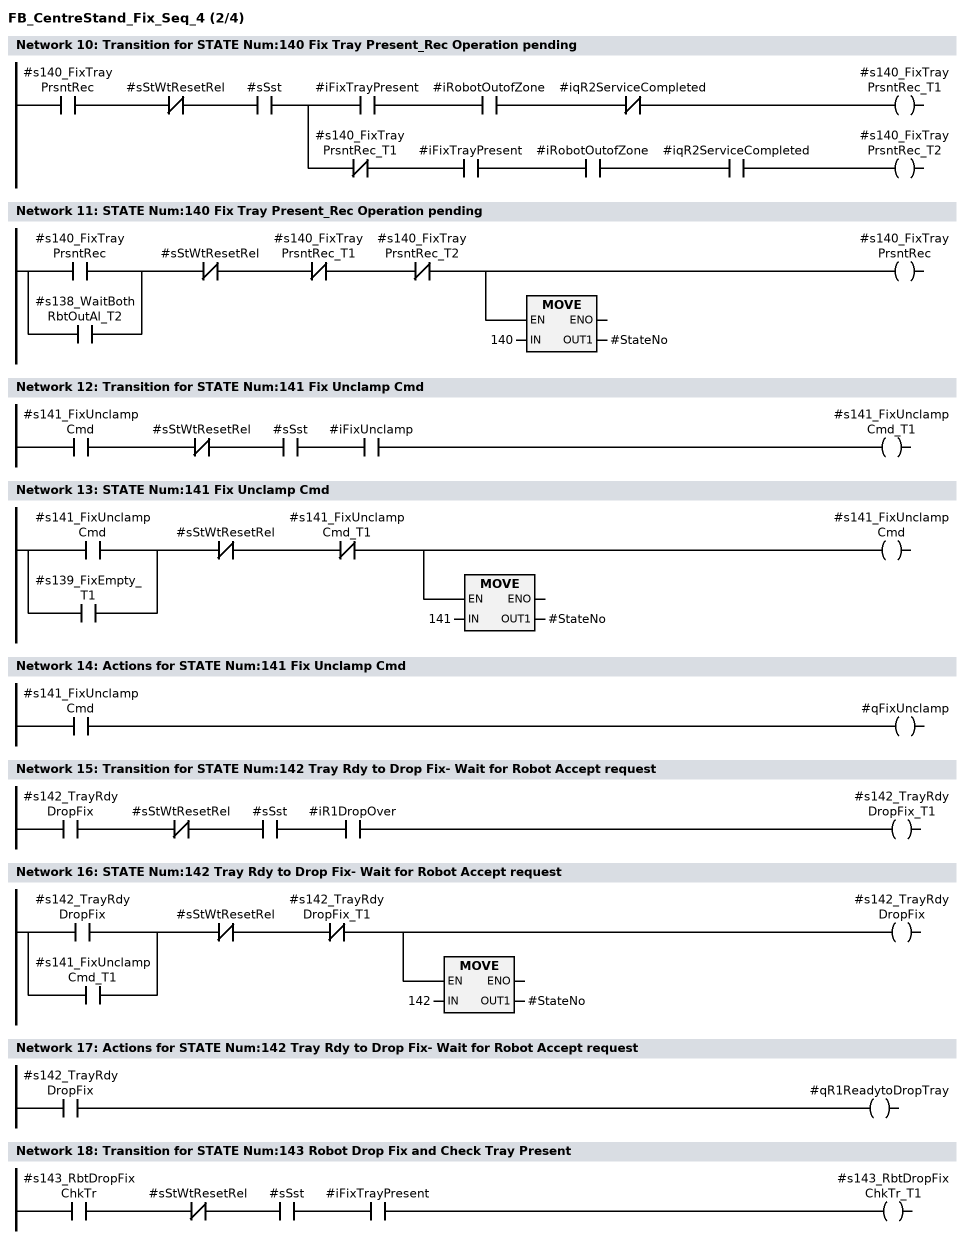
   RUNG wire#powerrail
      Contact( #s140_FixTrayPrsntRec )
      I_Contact( #sStWtResetRel )
      Contact( #sSst )
      wire#w1
      Contact( #iFixTrayPresent )
      Contact( #iRobotOutofZone )
      I_Contact( #iqR2ServiceCompleted )
      Coil( #s140_FixTrayPrsntRec_T1 )
   END_RUNG
   RUNG wire#w1
      I_Contact( #s140_FixTrayPrsntRec_T1 )
      Contact( #iFixTrayPresent )
      Contact( #iRobotOutofZone )
      Contact( #iqR2ServiceCompleted )
      Coil( #s140_FixTrayPrsntRec_T2 )
   END_RUNG
   // the same network as SCL:
   #_w1 := #s140_FixTrayPrsntRec AND NOT #sStWtResetRel AND #sSst;
   #s140_FixTrayPrsntRec_T1 := #_w1 AND #iFixTrayPresent AND #iRobotOutofZone AND NOT #iqR2ServiceCompleted;
   #s140_FixTrayPrsntRec_T2 := #_w1 AND NOT #s140_FixTrayPrsntRec_T1 AND #iFixTrayPresent AND #iRobotOutofZone AND #iqR2ServiceCompleted;
END_REGION

REGION Network 11: STATE Num:140 Fix Tray Present_Rec Operation pending
   RUNG wire#powerrail
      Contact( #s140_FixTrayPrsntRec )
      wire#w1
      I_Contact( #sStWtResetRel )
      I_Contact( #s140_FixTrayPrsntRec_T1 )
      I_Contact( #s140_FixTrayPrsntRec_T2 )
      wire#w2
      Coil( #s140_FixTrayPrsntRec )
   END_RUNG
   RUNG wire#powerrail
      Contact( #s138_WaitBothRbtOutAl_T2 )
   END_RUNG wire#w1
   RUNG wire#w2
      { S7_GenerateENO := "TRUE" } Move(in := 140, out1 => #StateNo)
   END_RUNG
   // the same network as SCL:
   #s140_FixTrayPrsntRec := (#s140_FixTrayPrsntRec OR #s138_WaitBothRbtOutAl_T2) AND NOT #sStWtResetRel AND NOT #s140_FixTrayPrsntRec_T1 AND NOT #s140_FixTrayPrsntRec_T2;
   IF #s140_FixTrayPrsntRec THEN #StateNo := 140; END_IF;
END_REGION

REGION Network 12: Transition for STATE Num:141 Fix Unclamp Cmd
   RUNG wire#powerrail
      Contact( #s141_FixUnclampCmd )
      I_Contact( #sStWtResetRel )
      Contact( #sSst )
      Contact( #iFixUnclamp )
      Coil( #s141_FixUnclampCmd_T1 )
   END_RUNG
   // the same network as SCL:
   #s141_FixUnclampCmd_T1 := #s141_FixUnclampCmd AND NOT #sStWtResetRel AND #sSst AND #iFixUnclamp;
END_REGION

REGION Network 13: STATE Num:141 Fix Unclamp Cmd
   RUNG wire#powerrail
      Contact( #s141_FixUnclampCmd )
      wire#w1
      I_Contact( #sStWtResetRel )
      I_Contact( #s141_FixUnclampCmd_T1 )
      wire#w2
      Coil( #s141_FixUnclampCmd )
   END_RUNG
   RUNG wire#powerrail
      Contact( #s139_FixEmpty_T1 )
   END_RUNG wire#w1
   RUNG wire#w2
      { S7_GenerateENO := "TRUE" } Move(in := 141, out1 => #StateNo)
   END_RUNG
   // the same network as SCL:
   #s141_FixUnclampCmd := (#s141_FixUnclampCmd OR #s139_FixEmpty_T1) AND NOT #sStWtResetRel AND NOT #s141_FixUnclampCmd_T1;
   IF #s141_FixUnclampCmd THEN #StateNo := 141; END_IF;
END_REGION

REGION Network 14: Actions for STATE Num:141 Fix Unclamp Cmd
   RUNG wire#powerrail
      Contact( #s141_FixUnclampCmd )
      Coil( #qFixUnclamp )
   END_RUNG
   // the same network as SCL:
   #qFixUnclamp := #s141_FixUnclampCmd;
END_REGION

REGION Network 15: Transition for STATE Num:142 Tray Rdy to Drop Fix- Wait for Robot Accept request
   RUNG wire#powerrail
      Contact( #s142_TrayRdyDropFix )
      I_Contact( #sStWtResetRel )
      Contact( #sSst )
      Contact( #iR1DropOver )
      Coil( #s142_TrayRdyDropFix_T1 )
   END_RUNG
   // the same network as SCL:
   #s142_TrayRdyDropFix_T1 := #s142_TrayRdyDropFix AND NOT #sStWtResetRel AND #sSst AND #iR1DropOver;
END_REGION

REGION Network 16: STATE Num:142 Tray Rdy to Drop Fix- Wait for Robot Accept request
   RUNG wire#powerrail
      Contact( #s142_TrayRdyDropFix )
      wire#w1
      I_Contact( #sStWtResetRel )
      I_Contact( #s142_TrayRdyDropFix_T1 )
      wire#w2
      Coil( #s142_TrayRdyDropFix )
   END_RUNG
   RUNG wire#powerrail
      Contact( #s141_FixUnclampCmd_T1 )
   END_RUNG wire#w1
   RUNG wire#w2
      { S7_GenerateENO := "TRUE" } Move(in := 142, out1 => #StateNo)
   END_RUNG
   // the same network as SCL:
   #s142_TrayRdyDropFix := (#s142_TrayRdyDropFix OR #s141_FixUnclampCmd_T1) AND NOT #sStWtResetRel AND NOT #s142_TrayRdyDropFix_T1;
   IF #s142_TrayRdyDropFix THEN #StateNo := 142; END_IF;
END_REGION

REGION Network 17: Actions for STATE Num:142 Tray Rdy to Drop Fix- Wait for Robot Accept request
   RUNG wire#powerrail
      Contact( #s142_TrayRdyDropFix )
      Coil( #qR1ReadytoDropTray )
   END_RUNG
   // the same network as SCL:
   #qR1ReadytoDropTray := #s142_TrayRdyDropFix;
END_REGION

REGION Network 18: Transition for STATE Num:143 Robot Drop Fix and Check Tray Present
   RUNG wire#powerrail
      Contact( #s143_RbtDropFixChkTr )
      I_Contact( #sStWtResetRel )
      Contact( #sSst )
      Contact( #iFixTrayPresent )
      Coil( #s143_RbtDropFixChkTr_T1 )
   END_RUNG
   // the same network as SCL:
   #s143_RbtDropFixChkTr_T1 := #s143_RbtDropFixChkTr AND NOT #sStWtResetRel AND #sSst AND #iFixTrayPresent;
END_REGION

REGION Network 19: STATE Num:143 Robot Drop Fix and Check Tray Present
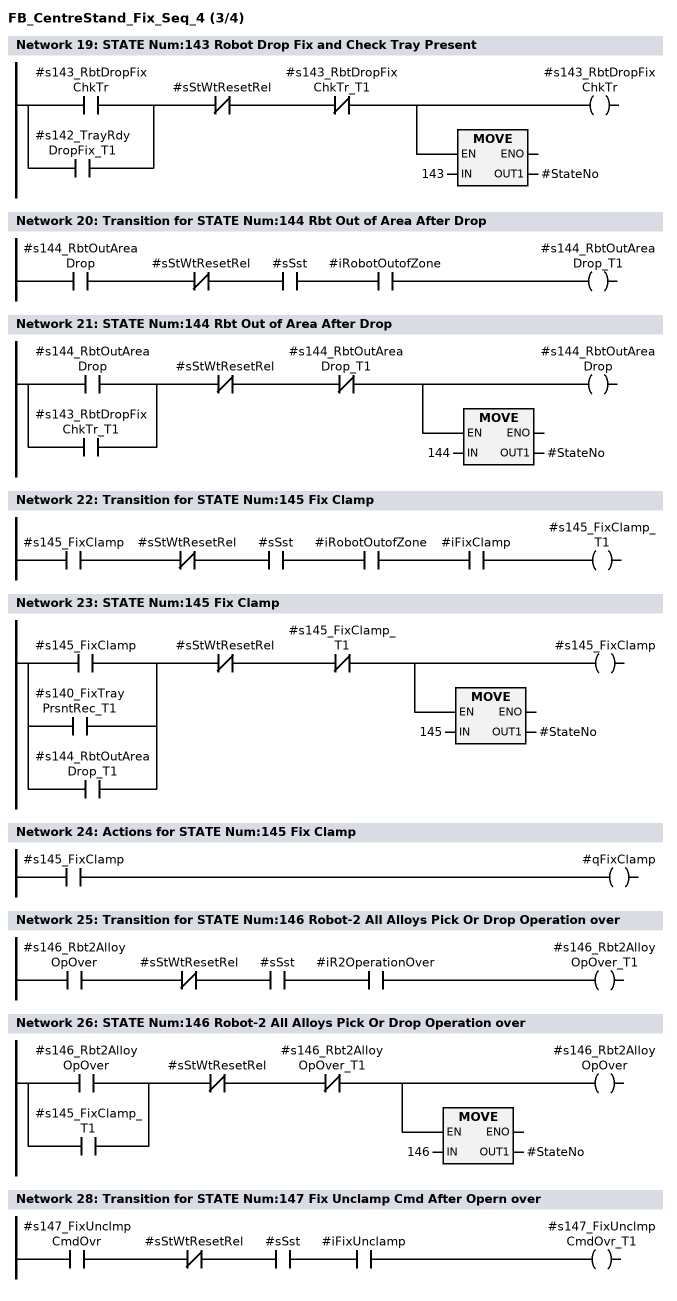
   RUNG wire#powerrail
      Contact( #s143_RbtDropFixChkTr )
      wire#w1
      I_Contact( #sStWtResetRel )
      I_Contact( #s143_RbtDropFixChkTr_T1 )
      wire#w2
      Coil( #s143_RbtDropFixChkTr )
   END_RUNG
   RUNG wire#powerrail
      Contact( #s142_TrayRdyDropFix_T1 )
   END_RUNG wire#w1
   RUNG wire#w2
      { S7_GenerateENO := "TRUE" } Move(in := 143, out1 => #StateNo)
   END_RUNG
   // the same network as SCL:
   #s143_RbtDropFixChkTr := (#s143_RbtDropFixChkTr OR #s142_TrayRdyDropFix_T1) AND NOT #sStWtResetRel AND NOT #s143_RbtDropFixChkTr_T1;
   IF #s143_RbtDropFixChkTr THEN #StateNo := 143; END_IF;
END_REGION

REGION Network 20: Transition for STATE Num:144 Rbt Out of Area After Drop
   RUNG wire#powerrail
      Contact( #s144_RbtOutAreaDrop )
      I_Contact( #sStWtResetRel )
      Contact( #sSst )
      Contact( #iRobotOutofZone )
      Coil( #s144_RbtOutAreaDrop_T1 )
   END_RUNG
   // the same network as SCL:
   #s144_RbtOutAreaDrop_T1 := #s144_RbtOutAreaDrop AND NOT #sStWtResetRel AND #sSst AND #iRobotOutofZone;
END_REGION

REGION Network 21: STATE Num:144 Rbt Out of Area After Drop
   RUNG wire#powerrail
      Contact( #s144_RbtOutAreaDrop )
      wire#w1
      I_Contact( #sStWtResetRel )
      I_Contact( #s144_RbtOutAreaDrop_T1 )
      wire#w2
      Coil( #s144_RbtOutAreaDrop )
   END_RUNG
   RUNG wire#powerrail
      Contact( #s143_RbtDropFixChkTr_T1 )
   END_RUNG wire#w1
   RUNG wire#w2
      { S7_GenerateENO := "TRUE" } Move(in := 144, out1 => #StateNo)
   END_RUNG
   // the same network as SCL:
   #s144_RbtOutAreaDrop := (#s144_RbtOutAreaDrop OR #s143_RbtDropFixChkTr_T1) AND NOT #sStWtResetRel AND NOT #s144_RbtOutAreaDrop_T1;
   IF #s144_RbtOutAreaDrop THEN #StateNo := 144; END_IF;
END_REGION

REGION Network 22: Transition for STATE Num:145 Fix Clamp
   RUNG wire#powerrail
      Contact( #s145_FixClamp )
      I_Contact( #sStWtResetRel )
      Contact( #sSst )
      Contact( #iRobotOutofZone )
      Contact( #iFixClamp )
      Coil( #s145_FixClamp_T1 )
   END_RUNG
   // the same network as SCL:
   #s145_FixClamp_T1 := #s145_FixClamp AND NOT #sStWtResetRel AND #sSst AND #iRobotOutofZone AND #iFixClamp;
END_REGION

REGION Network 23: STATE Num:145 Fix Clamp
   RUNG wire#powerrail
      Contact( #s145_FixClamp )
      wire#w1
      I_Contact( #sStWtResetRel )
      I_Contact( #s145_FixClamp_T1 )
      wire#w2
      Coil( #s145_FixClamp )
   END_RUNG
   RUNG wire#powerrail
      Contact( #s140_FixTrayPrsntRec_T1 )
   END_RUNG wire#w1
   RUNG wire#powerrail
      Contact( #s144_RbtOutAreaDrop_T1 )
   END_RUNG wire#w1
   RUNG wire#w2
      { S7_GenerateENO := "TRUE" } Move(in := 145, out1 => #StateNo)
   END_RUNG
   // the same network as SCL:
   #s145_FixClamp := (#s145_FixClamp OR #s140_FixTrayPrsntRec_T1 OR #s144_RbtOutAreaDrop_T1) AND NOT #sStWtResetRel AND NOT #s145_FixClamp_T1;
   IF #s145_FixClamp THEN #StateNo := 145; END_IF;
END_REGION

REGION Network 24: Actions for STATE Num:145 Fix Clamp
   RUNG wire#powerrail
      Contact( #s145_FixClamp )
      Coil( #qFixClamp )
   END_RUNG
   // the same network as SCL:
   #qFixClamp := #s145_FixClamp;
END_REGION

REGION Network 25: Transition for STATE Num:146 Robot-2 All Alloys Pick Or Drop Operation over
   RUNG wire#powerrail
      Contact( #s146_Rbt2AlloyOpOver )
      I_Contact( #sStWtResetRel )
      Contact( #sSst )
      Contact( #iR2OperationOver )
      Coil( #s146_Rbt2AlloyOpOver_T1 )
   END_RUNG
   // the same network as SCL:
   #s146_Rbt2AlloyOpOver_T1 := #s146_Rbt2AlloyOpOver AND NOT #sStWtResetRel AND #sSst AND #iR2OperationOver;
END_REGION

REGION Network 26: STATE Num:146 Robot-2 All Alloys Pick Or Drop Operation over
   RUNG wire#powerrail
      Contact( #s146_Rbt2AlloyOpOver )
      wire#w1
      I_Contact( #sStWtResetRel )
      I_Contact( #s146_Rbt2AlloyOpOver_T1 )
      wire#w2
      Coil( #s146_Rbt2AlloyOpOver )
   END_RUNG
   RUNG wire#powerrail
      Contact( #s145_FixClamp_T1 )
   END_RUNG wire#w1
   RUNG wire#w2
      { S7_GenerateENO := "TRUE" } Move(in := 146, out1 => #StateNo)
   END_RUNG
   // the same network as SCL:
   #s146_Rbt2AlloyOpOver := (#s146_Rbt2AlloyOpOver OR #s145_FixClamp_T1) AND NOT #sStWtResetRel AND NOT #s146_Rbt2AlloyOpOver_T1;
   IF #s146_Rbt2AlloyOpOver THEN #StateNo := 146; END_IF;
END_REGION

REGION Network 27 (STL): Actions for STATE Num:146 Robot-2 All Alloys Pick Or Drop Operation over
         A     #s146_Rbt2AlloyOpOver;
         =     #qR2OperationStart;
         A     #iR2ServiceActivated;
         S     #iqR2ServiceActive;
         A     #iR2OperationOver;
         A     #iqR2ServiceActive;
         R     #iqR2ServiceActive;
END_REGION

REGION Network 28: Transition for STATE Num:147 Fix Unclamp Cmd After Opern over
   RUNG wire#powerrail
      Contact( #s147_FixUnclmpCmdOvr )
      I_Contact( #sStWtResetRel )
      Contact( #sSst )
      Contact( #iFixUnclamp )
      Coil( #s147_FixUnclmpCmdOvr_T1 )
   END_RUNG
   // the same network as SCL:
   #s147_FixUnclmpCmdOvr_T1 := #s147_FixUnclmpCmdOvr AND NOT #sStWtResetRel AND #sSst AND #iFixUnclamp;
END_REGION

REGION Network 29: STATE Num:147 Fix Unclamp Cmd After Opern over
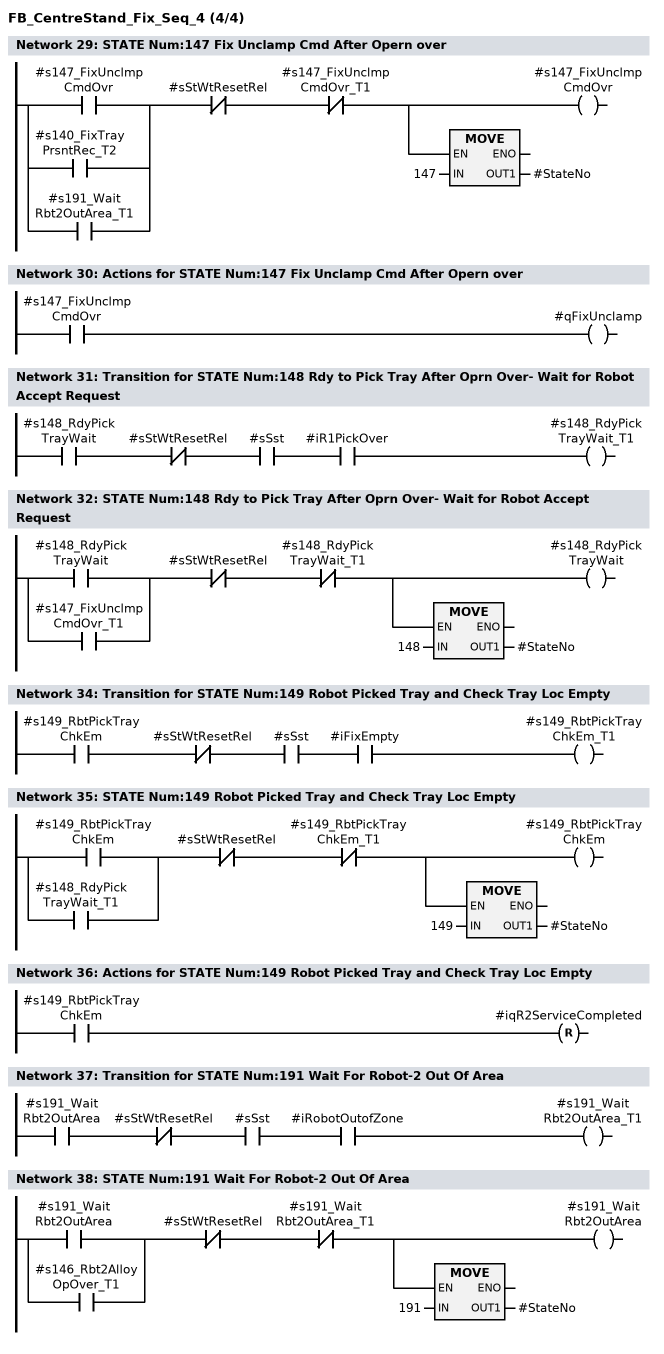
   RUNG wire#powerrail
      Contact( #s147_FixUnclmpCmdOvr )
      wire#w1
      I_Contact( #sStWtResetRel )
      I_Contact( #s147_FixUnclmpCmdOvr_T1 )
      wire#w2
      Coil( #s147_FixUnclmpCmdOvr )
   END_RUNG
   RUNG wire#powerrail
      Contact( #s140_FixTrayPrsntRec_T2 )
   END_RUNG wire#w1
   RUNG wire#powerrail
      Contact( #s191_WaitRbt2OutArea_T1 )
   END_RUNG wire#w1
   RUNG wire#w2
      { S7_GenerateENO := "TRUE" } Move(in := 147, out1 => #StateNo)
   END_RUNG
   // the same network as SCL:
   #s147_FixUnclmpCmdOvr := (#s147_FixUnclmpCmdOvr OR #s140_FixTrayPrsntRec_T2 OR #s191_WaitRbt2OutArea_T1) AND NOT #sStWtResetRel AND NOT #s147_FixUnclmpCmdOvr_T1;
   IF #s147_FixUnclmpCmdOvr THEN #StateNo := 147; END_IF;
END_REGION

REGION Network 30: Actions for STATE Num:147 Fix Unclamp Cmd After Opern over
   RUNG wire#powerrail
      Contact( #s147_FixUnclmpCmdOvr )
      Coil( #qFixUnclamp )
   END_RUNG
   // the same network as SCL:
   #qFixUnclamp := #s147_FixUnclmpCmdOvr;
END_REGION

REGION Network 31: Transition for STATE Num:148 Rdy to Pick Tray After Oprn Over- Wait for Robot Accept Request
   RUNG wire#powerrail
      Contact( #s148_RdyPickTrayWait )
      I_Contact( #sStWtResetRel )
      Contact( #sSst )
      Contact( #iR1PickOver )
      Coil( #s148_RdyPickTrayWait_T1 )
   END_RUNG
   // the same network as SCL:
   #s148_RdyPickTrayWait_T1 := #s148_RdyPickTrayWait AND NOT #sStWtResetRel AND #sSst AND #iR1PickOver;
END_REGION

REGION Network 32: STATE Num:148 Rdy to Pick Tray After Oprn Over- Wait for Robot Accept Request
   RUNG wire#powerrail
      Contact( #s148_RdyPickTrayWait )
      wire#w1
      I_Contact( #sStWtResetRel )
      I_Contact( #s148_RdyPickTrayWait_T1 )
      wire#w2
      Coil( #s148_RdyPickTrayWait )
   END_RUNG
   RUNG wire#powerrail
      Contact( #s147_FixUnclmpCmdOvr_T1 )
   END_RUNG wire#w1
   RUNG wire#w2
      { S7_GenerateENO := "TRUE" } Move(in := 148, out1 => #StateNo)
   END_RUNG
   // the same network as SCL:
   #s148_RdyPickTrayWait := (#s148_RdyPickTrayWait OR #s147_FixUnclmpCmdOvr_T1) AND NOT #sStWtResetRel AND NOT #s148_RdyPickTrayWait_T1;
   IF #s148_RdyPickTrayWait THEN #StateNo := 148; END_IF;
END_REGION

REGION Network 33 (STL): Actions for STATE Num:148 Rdy to Pick Tray After Oprn Over- Wait for Robot Accept Request
         A     #s148_RdyPickTrayWait;
         =     #qR1ReadytoPickTray;
         A     #iR1PickOver;
         R     #iqR2ServiceCompleted;
END_REGION

REGION Network 34: Transition for STATE Num:149 Robot Picked Tray and Check Tray Loc Empty
   RUNG wire#powerrail
      Contact( #s149_RbtPickTrayChkEm )
      I_Contact( #sStWtResetRel )
      Contact( #sSst )
      Contact( #iFixEmpty )
      Coil( #s149_RbtPickTrayChkEm_T1 )
   END_RUNG
   // the same network as SCL:
   #s149_RbtPickTrayChkEm_T1 := #s149_RbtPickTrayChkEm AND NOT #sStWtResetRel AND #sSst AND #iFixEmpty;
END_REGION

REGION Network 35: STATE Num:149 Robot Picked Tray and Check Tray Loc Empty
   RUNG wire#powerrail
      Contact( #s149_RbtPickTrayChkEm )
      wire#w1
      I_Contact( #sStWtResetRel )
      I_Contact( #s149_RbtPickTrayChkEm_T1 )
      wire#w2
      Coil( #s149_RbtPickTrayChkEm )
   END_RUNG
   RUNG wire#powerrail
      Contact( #s148_RdyPickTrayWait_T1 )
   END_RUNG wire#w1
   RUNG wire#w2
      { S7_GenerateENO := "TRUE" } Move(in := 149, out1 => #StateNo)
   END_RUNG
   // the same network as SCL:
   #s149_RbtPickTrayChkEm := (#s149_RbtPickTrayChkEm OR #s148_RdyPickTrayWait_T1) AND NOT #sStWtResetRel AND NOT #s149_RbtPickTrayChkEm_T1;
   IF #s149_RbtPickTrayChkEm THEN #StateNo := 149; END_IF;
END_REGION

REGION Network 36: Actions for STATE Num:149 Robot Picked Tray and Check Tray Loc Empty
   RUNG wire#powerrail
      Contact( #s149_RbtPickTrayChkEm )
      R_Coil( #iqR2ServiceCompleted )
   END_RUNG
   // the same network as SCL:
   IF #s149_RbtPickTrayChkEm THEN #iqR2ServiceCompleted := FALSE; END_IF;
END_REGION

REGION Network 37: Transition for STATE Num:191 Wait For Robot-2 Out Of Area
   RUNG wire#powerrail
      Contact( #s191_WaitRbt2OutArea )
      I_Contact( #sStWtResetRel )
      Contact( #sSst )
      Contact( #iRobotOutofZone )
      Coil( #s191_WaitRbt2OutArea_T1 )
   END_RUNG
   // the same network as SCL:
   #s191_WaitRbt2OutArea_T1 := #s191_WaitRbt2OutArea AND NOT #sStWtResetRel AND #sSst AND #iRobotOutofZone;
END_REGION

REGION Network 38: STATE Num:191 Wait For Robot-2 Out Of Area
   RUNG wire#powerrail
      Contact( #s191_WaitRbt2OutArea )
      wire#w1
      I_Contact( #sStWtResetRel )
      I_Contact( #s191_WaitRbt2OutArea_T1 )
      wire#w2
      Coil( #s191_WaitRbt2OutArea )
   END_RUNG
   RUNG wire#powerrail
      Contact( #s146_Rbt2AlloyOpOver_T1 )
   END_RUNG wire#w1
   RUNG wire#w2
      { S7_GenerateENO := "TRUE" } Move(in := 191, out1 => #StateNo)
   END_RUNG
   // the same network as SCL:
   #s191_WaitRbt2OutArea := (#s191_WaitRbt2OutArea OR #s146_Rbt2AlloyOpOver_T1) AND NOT #sStWtResetRel AND NOT #s191_WaitRbt2OutArea_T1;
   IF #s191_WaitRbt2OutArea THEN #StateNo := 191; END_IF;
END_REGION
END_FUNCTION_BLOCK

